/// Read a server log of the RC line by line into LogFile
FUNCTION_BLOCK MC_ReadServerLogFB EXTENDS RobotLibraryBaseExecuteFB
// -------------------------------------------------------------------------
//  SRCI Robot Library
// -------------------------------------------------------------------------
//
//  Object:      MC_ReadServerLogFB
//  Author:      Thorsten Brach
//  Date:        2026-10-23
//
//  Description:
//    ReadServerLog (spec 6.2.6, type 9004): reads the server log ParCmd.ServerLogID from
//    ParCmd.StartLine on into the array LogFile, one CSV line per element. The RC sends a log line in
//    parts of up to 179 characters; the block joins them. The transfer ends with Done when the RC
//    reports the end of the log or when LogFile is full. A rising edge of Execute during the transfer
//    starts it again.
//    Telegram layout of SRCI SDK 1.1.2 (Offset as request counter, IsStartOfLine / IsEndOfLine /
//    EndOfLogReached / LogLine in the response); spec table 6-123 / 6-124 differ.
//
//  Copyright:
//    (C) 2026 Thorsten Brach. All rights reserved
//             Licensed under the MIT License.
//
//  Disclaimer:
//    This project is provided without any guarantee and can be used for
//    private and commercial purposes. Any use is at the user's
//    own risk and responsibility.
//
// -------------------------------------------------------------------------
VAR_INPUT
  /// command parameter
  ParCmd          : ReadServerLogParCmd;
END_VAR
VAR_OUTPUT
  /// Command is transferred and confirmed by the RC
  CommandBuffered : BOOL;
  /// command outputs
  OutCmd          : ReadServerLogOutCmd;
END_VAR
VAR_IN_OUT
  /// Requested log file: one log line per element
  LogFile         : ARRAY [*] OF STRING(RobotLibraryParameter.LOG_LINE_LEN);
END_VAR
VAR
  /// internal copy of command parameter
 _parCmd          : ReadServerLogParCmd;
  /// command data to send
 _command         : ReadServerLogSendData;
  /// response data received
 _response        : ReadServerLogRecvData;
  /// a part of the log was received and must be stored in LogFile (StoreLogContent)
 _contentReceived : BOOL;
  /// the response to the current Offset was handled
 _offsetHandled   : BOOL;
  /// new rising edge of Execute during the transfer: start again after the end of this one
 _restart         : BOOL;
  /// index of the element of LogFile for the current log line
 _line            : DINT;
  /// number of elements of LogFile used by this transfer
 _lines           : DINT;
  /// a log line is open (parts received, end of line not yet)
 _lineOpen        : BOOL;
  /// characters of the current log line
 _lineLen         : DINT;
  /// characters copied from the received part
 _copyLen         : DINT;
END_VAR

            SUPER^(AxesGroup := AxesGroup);

// store the received part of the log (LogFile is only reachable in the call of the block)
StoreLogContent( AxesGroup := AxesGroup, LogFile := LogFile );
          

METHOD INTERNAL CheckAddParameter : BOOL
VAR_INPUT
  /// Payload pointer
  PayloadPtr : UDINT;
END_VAR
VAR
  /// Payload as byte array
  Payload    : ARRAY [1..SIZEOF(_command)] OF BYTE;
  /// Null Byte array
  Null       : ARRAY [1..SIZEOF(_command)] OF BYTE;
  /// Data length to compare
  DataLen    : UDINT;
END_VAR
                  // Payload pointer must be decreased by one byte, because ADR(Payload) is already one byte !
PayloadPtr := LIMIT (0, PayloadPtr - 1, SIZEOF(Payload) -1);
// Convert command struct to payload array
SysDepMemCpy( pDest := ADR(Payload), pSrc := ADR(_command), DataLen := SIZEOF(_command));
// Calculate the data length to compare - at least one byte must be compared !
DataLen := LIMIT(1, SIZEOF(Payload) - PayloadPtr, SIZEOF(Payload));
// Compare Payload-Array with Null-Byte-Array
CheckAddParameter := SysDepMemCmp( pData1 := ADR(Payload) + PayloadPtr , pData2 := ADR(Null), DataLen := DataLen) <>  RobotLibraryConstants.OK ;
                
END_METHOD

METHOD PROTECTED CheckFunctionSupported : BOOL
VAR_IN_OUT
  /// Robot assignment of function
  AxesGroup : AxesGroup;
END_VAR
                  // ReadServerLog is a mandatory function of the profile Core (spec table 6-119): the RC
// reports no bit for it in RCSupportedFunctions
CheckFunctionSupported := TRUE;
                
END_METHOD

METHOD PROTECTED CheckParameterChanged : BOOL
VAR_IN_OUT
  /// Robot assignment of function
  AxesGroup    : AxesGroup;
END_VAR
                  // The parameters of the transfer are taken with the rising edge of Execute; during the transfer
// only the block itself sends updates (next part of the log: Offset, end: Enable FALSE)
IF ( _stepCmd = 0 )
THEN
  RETURN;
END_IF

IF ( _parameterUpdateInternal )
THEN
  // reset internal flag for send parameter update
 _parameterUpdateInternal := FALSE;
  // inc parameter sequence
 _command.ParSeq := _command.ParSeq + 1;
  // update command data
  CommandData := CreateCommandPayload(AxesGroup := AxesGroup); // ( Access via reference to rCommandFB in ACR )
  // notify active command register
  AxesGroup.Acyclic.ActiveCommandRegister.NotifyParameterChanged := _uniqueID;
END_IF
                
END_METHOD

METHOD PROTECTED CheckParameterValid : BOOL
VAR_IN_OUT
  /// Robot assignment of function
  AxesGroup : AxesGroup;
END_VAR
                  CheckParameterValid := TRUE;

// Check ParCmd.ExportMode: only 0 (output LogFile), the export to a file is optional (table 6-119)
IF ( ParCmd.ExportMode <> 0 )
THEN
  // Parameter not valid
  CheckParameterValid := FALSE;
  // Set error
  SetError( ErrorID := RobotLibraryErrorIdEnum.ERR_EXPORTMODE_NOT_EXIST, Overwrite := TRUE );
  // Create log entry
  CreateLogMessagePara1 ( Timestamp   := AxesGroup.State.SystemTime,
                          MessageType := MessageType.CMD,
                          Severity    := Severity.ERROR,
                          MessageCode := ErrorID,
                          MessageText := 'Invalid Parameter ParCmd.ExportMode = {1}',
                          Para1       := USINT_TO_STRING(ParCmd.ExportMode));
  RETURN;
END_IF

// Check ParCmd.StartLine: the first line is 1 (log header)
IF ( ParCmd.StartLine = 0 )
THEN
  // Parameter not valid
  CheckParameterValid := FALSE;
  // Set error
  SetError( ErrorID := RobotLibraryErrorIdEnum.ERR_INVALID_PAR_CMD, Overwrite := TRUE );
  // Create log entry
  CreateLogMessagePara1 ( Timestamp   := AxesGroup.State.SystemTime,
                          MessageType := MessageType.CMD,
                          Severity    := Severity.ERROR,
                          MessageCode := ErrorID,
                          MessageText := 'Invalid Parameter ParCmd.StartLine = {1}',
                          Para1       := UDINT_TO_STRING(ParCmd.StartLine));
  RETURN;
END_IF

// Check ParCmd.ServerLogID: -1 (latest), 0 (oldest) or an ID
IF ( ParCmd.ServerLogID < -1 )
THEN
  // Parameter not valid
  CheckParameterValid := FALSE;
  // Set error
  SetError( ErrorID := RobotLibraryErrorIdEnum.ERR_INVALID_PAR_CMD, Overwrite := TRUE );
  // Create log entry
  CreateLogMessagePara1 ( Timestamp   := AxesGroup.State.SystemTime,
                          MessageType := MessageType.CMD,
                          Severity    := Severity.ERROR,
                          MessageCode := ErrorID,
                          MessageText := 'Invalid Parameter ParCmd.ServerLogID = {1}',
                          Para1       := INT_TO_STRING(ParCmd.ServerLogID));
  RETURN;
END_IF
                
END_METHOD

METHOD INTERNAL CreateCommandPayload : RobotLibraryCommandDataFB
VAR_IN_OUT
  /// Robot assignment of function
  AxesGroup : AxesGroup;
END_VAR
VAR
  /// internal index for loops
 _idx          : DINT;
  /// Parameter count
 _parameterCnt : DINT;
END_VAR
// Sent CMD payload (PLC to RC) of "ReadServerLog" - layout of SRCI SDK 1.1.2 (spec table 6-123
// has no Offset, ContextFilter at byte 12)
// --------------------------
// Header
// --------------------------
// Byte 00 : UINT  - Type HB
// Byte 01 :       - Type LB
// Byte 02 : USINT - Reserve | ExecutionMode
// Byte 03 : USINT - ParSeq  | Priority
// --------------------------
// Datablock
// --------------------------
// Byte 04 : BYTE  - Bit 0: Enable
// Byte 05 : BYTE  - Reserved
// Byte 06 : UINT  - ServerLogID HB
// Byte 07 :       - ServerLogID LB
// Byte 08 : UDINT - StartLine
// Byte 12 : UDINT - Offset
// Byte 16 : USINT - ContextFilter[0]
// ...
// Byte 25 : USINT - ContextFilter[9]
// --------------------------
                  // set command parameter
_command.CmdTyp      :=  CmdType.ReadServerLog;
// spec table 6-121: parallel only (default of ExecMode, FB_init)
_command.ExecMode    :=  ExecMode;
_command.ParSeq      := _command.ParSeq;
_command.Priority    :=  Priority;
_command.Reserve     := 0;
// -1 (latest) -> 16#FFFF
_command.ServerLogID := INT_TO_UINT(_parCmd.ServerLogID);
_command.StartLine   := _parCmd.StartLine;
FOR _idx := 0 TO 9
DO
  _command.ContextFilter[_idx] := _parCmd.ContextFilter[_idx];
END_FOR

// copy command data to header
_cmdHeader := _command;
// call base implementation to copy header to payload buffer
CreateCommandPayload := SUPER^.CreateCommandPayload(AxesGroup := AxesGroup);

// Check parameter must be added ?
IF ( CheckAddParameter(CreateCommandPayload.PayloadPtr))
THEN
  // add command.Enable
  CreateCommandPayload.AddBool(_command.Enable);
  // inc parameter counter
 _parameterCnt := _parameterCnt + 1;
END_IF

// Check parameter must be added ?
IF ( CheckAddParameter(CreateCommandPayload.PayloadPtr))
THEN
  // add command.Reserve
  CreateCommandPayload.AddByte(_command.Reserve);
  // inc parameter counter
 _parameterCnt := _parameterCnt + 1;
END_IF

// Check parameter must be added ?
IF ( CheckAddParameter(CreateCommandPayload.PayloadPtr))
THEN
  // add command.ServerLogID
  CreateCommandPayload.AddUint(_command.ServerLogID);
  // inc parameter counter
 _parameterCnt := _parameterCnt + 1;
END_IF

// Check parameter must be added ?
IF ( CheckAddParameter(CreateCommandPayload.PayloadPtr))
THEN
  // add command.StartLine
  CreateCommandPayload.AddUdint(_command.StartLine);
  // inc parameter counter
 _parameterCnt := _parameterCnt + 1;
END_IF

// Check parameter must be added ?
IF ( CheckAddParameter(CreateCommandPayload.PayloadPtr))
THEN
  // add command.Offset
  CreateCommandPayload.AddUdint(_command.Offset);
  // inc parameter counter
 _parameterCnt := _parameterCnt + 1;
END_IF

FOR _idx := 0 TO 9
DO
  // Check parameter must be added ?
  IF ( CheckAddParameter(CreateCommandPayload.PayloadPtr))
  THEN
    // add command.ContextFilter[x]
    CreateCommandPayload.AddUsint(_command.ContextFilter[_idx]);
    // inc parameter counter
   _parameterCnt := _parameterCnt + 1;
  END_IF
END_FOR

// Create logging
CreateCommandPayloadLog(AxesGroup := AxesGroup, ParameterCnt := _parameterCnt);
                
END_METHOD

METHOD INTERNAL CreateCommandPayloadLog
VAR_IN_OUT
  /// Robot assignment of function
  AxesGroup : AxesGroup;
END_VAR
VAR_INPUT
  /// Parameter count
  ParameterCnt : DINT;
END_VAR
VAR
  /// internal index for loops
 _idx : DINT;
END_VAR
                  // Create log entry for Parameter start
CreateLogMessagePara1 ( Timestamp   := AxesGroup.State.SystemTime,
                        MessageType := MessageType.CMD,
                        Severity    := Severity.DEBUG,
                        MessageCode := 0,
                        MessageText := 'Create command payload with {1} parameter(s) :',
                        Para1       := DINT_TO_STRING(ParameterCnt));

// Return if no parameter is remaining...
IF ( ParameterCnt = 0 ) THEN RETURN; END_IF
// dec remaining parameter(s)
ParameterCnt := ParameterCnt - 1;
// Create log entry for Command.Enable
CreateLogMessagePara1 ( Timestamp   := AxesGroup.State.SystemTime,
                        MessageType := MessageType.CMD,
                        Severity    := Severity.DEBUG,
                        MessageCode := 0,
                        MessageText := 'Command.Enable = {1}',
                        Para1       :=  BOOL_TO_STRING(_command.Enable));

// Return if no parameter is remaining...
IF ( ParameterCnt = 0 ) THEN RETURN; END_IF
// dec remaining parameter(s)
ParameterCnt := ParameterCnt - 1;
// Create log entry for Command.Reserve
CreateLogMessagePara1 ( Timestamp   := AxesGroup.State.SystemTime,
                        MessageType := MessageType.CMD,
                        Severity    := Severity.DEBUG,
                        MessageCode := 0,
                        MessageText := 'Command.Reserve = {1}',
                        Para1       :=  BYTE_TO_STRING(_command.Reserve));

// Return if no parameter is remaining...
IF ( ParameterCnt = 0 ) THEN RETURN; END_IF
// dec remaining parameter(s)
ParameterCnt := ParameterCnt - 1;
// Create log entry for Command.ServerLogID
CreateLogMessagePara1 ( Timestamp   := AxesGroup.State.SystemTime,
                        MessageType := MessageType.CMD,
                        Severity    := Severity.DEBUG,
                        MessageCode := 0,
                        MessageText := 'Command.ServerLogID = {1}',
                        Para1       :=  UINT_TO_STRING(_command.ServerLogID));

// Return if no parameter is remaining...
IF ( ParameterCnt = 0 ) THEN RETURN; END_IF
// dec remaining parameter(s)
ParameterCnt := ParameterCnt - 1;
// Create log entry for Command.StartLine
CreateLogMessagePara1 ( Timestamp   := AxesGroup.State.SystemTime,
                        MessageType := MessageType.CMD,
                        Severity    := Severity.DEBUG,
                        MessageCode := 0,
                        MessageText := 'Command.StartLine = {1}',
                        Para1       :=  UDINT_TO_STRING(_command.StartLine));

// Return if no parameter is remaining...
IF ( ParameterCnt = 0 ) THEN RETURN; END_IF
// dec remaining parameter(s)
ParameterCnt := ParameterCnt - 1;
// Create log entry for Command.Offset
CreateLogMessagePara1 ( Timestamp   := AxesGroup.State.SystemTime,
                        MessageType := MessageType.CMD,
                        Severity    := Severity.DEBUG,
                        MessageCode := 0,
                        MessageText := 'Command.Offset = {1}',
                        Para1       :=  UDINT_TO_STRING(_command.Offset));

FOR _idx := 0 TO 9
DO
  // Return if no parameter is remaining...
  IF ( ParameterCnt = 0 ) THEN RETURN; END_IF
  // dec remaining parameter(s)
  ParameterCnt := ParameterCnt - 1;
  // Create log entry for Command.ContextFilter
  CreateLogMessagePara2 ( Timestamp   := AxesGroup.State.SystemTime,
                          MessageType := MessageType.CMD,
                          Severity    := Severity.DEBUG,
                          MessageCode := 0,
                          MessageText := 'Command.ContextFilter[{2}] = {1}',
                          Para1       :=  USINT_TO_STRING(_command.ContextFilter[_idx]),
                          Para2       :=  DINT_TO_STRING(_idx));
END_FOR
                
END_METHOD

METHOD FB_init : BOOL
VAR_INPUT
  /// if TRUE, the retain variables are initialized (warm start / cold start)
  bInitRetains : BOOL;
  /// if TRUE, the instance afterwards gets moved into the copy code (online change)
  bInCopyCode  : BOOL;
END_VAR
                  MyType := 'MC_ReadServerLogFB';

// spec 6.2.6: processed with low priority because of its processing time
ExecMode := ExecutionMode.PARALLEL;
Priority := PriorityLevel.LOW;
                
END_METHOD

METHOD PROTECTED OnApplyOutCmd
VAR_INPUT
  /// Command message state
  State : CmdMessageState;
END_VAR
                  IF ( State = CmdMessageState.EMPTY )
THEN
  // Reset command outputs
  SysDepMemSet(pDest := ADR(OutCmd), Value := 0, DataLen := SIZEOF(OutCmd));
END_IF

// the counters of the log come with every part (StoreLogContent), the received lines are counted there
                
END_METHOD

METHOD PROTECTED OnExecRun : DINT
VAR_IN_OUT
  /// Robot assignment of function
  AxesGroup : AxesGroup;
END_VAR
                  // call base implementation
SUPER^.OnExecRun(AxesGroup := AxesGroup);

CASE _stepCmd OF

  00:  IF (( _execute_R.Q ) OR ( _restart )) AND ( NOT Error )
       THEN
        _restart := FALSE;
         // Check function is supported and parameter are valid ?
         IF (( CheckFunctionSupported( AxesGroup := AxesGroup )) AND
             ( CheckParameterValid   ( AxesGroup := AxesGroup )))
         THEN
           // set busy flag
           Busy := TRUE;
           // Reset command outputs
           SysDepMemSet(pDest := ADR(OutCmd), Value := 0, DataLen := SIZEOF(OutCmd));
           // apply command parameter
          _parCmd := ParCmd;
           // first element of LogFile, no open line
          _line            := 0;
          _lines           := 0;
          _lineOpen        := FALSE;
          _lineLen         := 0;
          _contentReceived := FALSE;
          _offsetHandled   := FALSE;
           // transfer on, first request
          _command.Enable := TRUE;
          _command.Offset := 1;
           // init parameter sequence
          _command.ParSeq := 1;
           // create command data
           CommandData := CreateCommandPayload(AxesGroup := AxesGroup);
           // Add command to active command register
          _uniqueID := AxesGroup.Acyclic.ActiveCommandRegister.AddCmd( pCommandFB := ADR(THIS^ ));
           // set timeout
           SetTimeout(PT := _timeoutCmd, rTimer := _timerCmd);
           // inc step counter
          _stepCmd := _stepCmd + 1;
         END_IF
       END_IF

  01:  // spec 6.2.6: a new rising edge of Execute during the transfer aborts it and starts the
       // command again. SRCI SDK 1.1 keeps the read position of a running command, so the transfer
       // ends first (Enable FALSE) and the command is added again (new ACR entry).
       IF ( _executeRestart_R.Q ) AND ( NOT _restart )
       THEN
        _restart := TRUE;
        _command.Enable := FALSE;
        _parameterUpdateInternal := TRUE;
       END_IF

       // Wait for responce received
       IF ( _responseReceived )
       THEN
         // reset response received flag
        _responseReceived := FALSE;

         CASE _response.State OF
           CmdMessageState.DONE:
             IF ( _restart )
             THEN
               // the old transfer ended: start again (step 00)
               Reset();
              _restart := TRUE;
             ELSE
               OnUpdateStateFlags(_response.State);
               // set timeout
               SetTimeout(PT := _timeoutCmd, rTimer := _timerCmd);
               // inc step counter
              _stepCmd := _stepCmd + 1;
             END_IF

           CmdMessageState.ABORTED, CmdMessageState.ERROR:
            _restart := FALSE;
             OnUpdateStateFlags(_response.State);
             // set timeout
             SetTimeout(PT := _timeoutCmd, rTimer := _timerCmd);
             // inc step counter
            _stepCmd := _stepCmd + 1;

         ELSE
           OnUpdateStateFlags(_response.State);
           // a part of the log for the current request ? (responses to older requests are ignored)
           IF (( _command.Enable                     ) AND
               ( NOT _restart                        ) AND
               ( NOT _offsetHandled                  ) AND
               ( _response.Offset = _command.Offset  ))
           THEN
            _offsetHandled   := TRUE;
            _contentReceived := TRUE;
           END_IF
         END_CASE
       END_IF

  02: IF ( NOT Execute)
      THEN
        Reset();
      END_IF

ELSE
  // invalid step
  SetError( ErrorID := RobotLibraryErrorIdEnum.ERR_INVALID_STEP, Overwrite := TRUE );
END_CASE

// Reset FB
IF ( NOT Execute ) AND ( NOT _restart )
THEN
  Reset();
END_IF
                
END_METHOD

METHOD PROTECTED OnUpdateStateFlags
VAR_INPUT
  /// Command message state
  State : CmdMessageState;
END_VAR
                  // Reset State flags
Done := FALSE;

CASE State OF
  // No operation or process is active
  CmdMessageState.EMPTY               :;
  // Created but not yet started
  CmdMessageState.CREATED             :;
  // Buffered and awaiting execution
  CmdMessageState.BUFFERED            : CommandBuffered := TRUE;
  // Buffered in planner for future execution
  CmdMessageState.BUFFERED_IN_PLANNER : CommandBuffered := TRUE;
  // Currently active and in progress
  CmdMessageState.ACTIVE              : CommandBuffered := TRUE;
  // Interrupted and awaiting continuation
  CmdMessageState.INTERRUPTED         :;
  // Requested for abort
  CmdMessageState.ABORT_REQUEST       :;
  // Successfully completed
  CmdMessageState.DONE                : Done            := TRUE;
                                        Busy            := FALSE;
  // Aborted before completion
  CmdMessageState.ABORTED             : Busy            := FALSE;
  // Encountered an error during execution
  CmdMessageState.ERROR               : Error           := TRUE;
                                        Busy            := FALSE;
END_CASE
                
END_METHOD

METHOD INTERNAL ParseResponsePayload : DINT
VAR_INPUT
  /// Response data
  ResponseData : RobotLibraryResponseDataFB;
  /// Timestamp
  Timestamp    : SystemTime;
END_VAR
VAR
  /// Parameter count
 _parameterCnt : DINT;
  /// Byte 13: line flags
 _flags        : BYTE;
END_VAR
// Received CMD payload (RC to PLC) of "ReadServerLog" - layout of SRCI SDK 1.1.2 (spec table
// 6-124: byte 13 only IsSplitLine, LogContent from byte 14)
// --------------------------
// Header
// --------------------------
// Byte 00 : USINT   - ParSeq | State
// Byte 01 : SINT    - AlarmMessageSeverity
// Byte 02 : UINT    - AlarmMessageCode HB
// Byte 03 :         - AlarmMessageCode LB
// --------------------------
// Datablock
// --------------------------
// Byte 04 : UDINT   - AvailableLogLines
// Byte 08 : UDINT   - AvailableFilteredLogLines
// Byte 12 : USINT   - LogContentLength
// Byte 13 : BYTE    - Bit 0: IsStartOfLine, Bit 1: IsEndOfLine, Bit 2: EndOfLogReached
// Byte 14 : UDINT   - LogLine
// Byte 18 : UDINT   - Offset
// Byte 22 : CHAR    - LogContent[0]
// ...
// Byte 200: CHAR    - LogContent[178]
// --------------------------
                  // call base implementation to parse the header from payload buffer
ResponseData.PayloadPtr := SUPER^.ParseResponsePayload(ResponseData := ResponseData, Timestamp := Timestamp);

// missing (trailing zero) bytes of the payload are 0, no values of the previous response
SysDepMemSet( pDest := ADR(_response), Value := 0, DataLen := SIZEOF(_response));

// copy parsed header to response
_response.ParSeq               := _rspHeader.ParSeq;
_response.State                := _rspHeader.State;
_response.AlarmMessageSeverity := _rspHeader.AlarmMessageSeverity;
_response.AlarmMessageCode     := _rspHeader.AlarmMessageCode;

// Check payload remaining ?
IF ( ResponseData.IsPayloadRemaining)
THEN
  // Get Response.AvailableLogLines
 _response.AvailableLogLines := ResponseData.GetUdint();
  // inc parameter counter
 _parameterCnt := _parameterCnt + 1;
END_IF

// Check payload remaining ?
IF ( ResponseData.IsPayloadRemaining)
THEN
  // Get Response.AvailableFilteredLogLines
 _response.AvailableFilteredLogLines := ResponseData.GetUdint();
  // inc parameter counter
 _parameterCnt := _parameterCnt + 1;
END_IF

// Check payload remaining ?
IF ( ResponseData.IsPayloadRemaining)
THEN
  // Get Response.LogContentLength
 _response.LogContentLength := ResponseData.GetUsint();
  // inc parameter counter
 _parameterCnt := _parameterCnt + 1;
END_IF

// Check payload remaining ?
IF ( ResponseData.IsPayloadRemaining)
THEN
  // Get Response.IsStartOfLine / IsEndOfLine / EndOfLogReached
 _flags                     := ResponseData.GetByte();
 _response.IsStartOfLine    := _flags.0;
 _response.IsEndOfLine      := _flags.1;
 _response.EndOfLogReached  := _flags.2;
  // inc parameter counter
 _parameterCnt := _parameterCnt + 1;
END_IF

// Check payload remaining ?
IF ( ResponseData.IsPayloadRemaining)
THEN
  // Get Response.LogLine
 _response.LogLine := ResponseData.GetUdint();
  // inc parameter counter
 _parameterCnt := _parameterCnt + 1;
END_IF

// Check payload remaining ?
IF ( ResponseData.IsPayloadRemaining)
THEN
  // Get Response.Offset
 _response.Offset := ResponseData.GetUdint();
  // inc parameter counter
 _parameterCnt := _parameterCnt + 1;
END_IF

// Check payload remaining ?
IF ( ResponseData.IsPayloadRemaining ) AND ( _response.LogContentLength > 0 )
THEN
  // Get Response.LogContent (LogContentLength characters)
 _response.LogContent := ResponseData.GetString( Size := MIN( USINT_TO_DINT(_response.LogContentLength), RobotLibraryConstants.SERVER_LOG_CONTENT_MAX ));
  // inc parameter counter
 _parameterCnt := _parameterCnt + 1;
END_IF

// Create logging
ParseResponsePayloadLog(ResponseData := ResponseData, Timestamp := Timestamp, ParameterCnt := _parameterCnt);
                
END_METHOD

METHOD INTERNAL ParseResponsePayloadLog
VAR_INPUT
  /// Response data
  ResponseData : RobotLibraryResponseDataFB;
  /// Timestamp
  Timestamp    : SystemTime;
  /// Parameter count
  ParameterCnt : DINT;
END_VAR
                  // Create log entry for Parameter start
CreateLogMessagePara1 ( Timestamp   := Timestamp,
                        MessageType := MessageType.CMD,
                        Severity    := Severity.DEBUG,
                        MessageCode := 0,
                        MessageText := '{1} parameter(s) to parse from the response data:',
                        Para1       := DINT_TO_STRING(ParameterCnt));

// Return if no parameter is remaining...
IF ( ParameterCnt = 0 ) THEN RETURN; END_IF
// dec remaining parameter(s)
ParameterCnt := ParameterCnt - 1;
// Create log entry for AvailableLogLines
CreateLogMessagePara1 ( Timestamp   := Timestamp,
                        MessageType := MessageType.CMD,
                        Severity    := Severity.DEBUG,
                        MessageCode := 0,
                        MessageText := 'Response.AvailableLogLines = {1}',
                        Para1       :=  UDINT_TO_STRING(_response.AvailableLogLines));

// Return if no parameter is remaining...
IF ( ParameterCnt = 0 ) THEN RETURN; END_IF
// dec remaining parameter(s)
ParameterCnt := ParameterCnt - 1;
// Create log entry for AvailableFilteredLogLines
CreateLogMessagePara1 ( Timestamp   := Timestamp,
                        MessageType := MessageType.CMD,
                        Severity    := Severity.DEBUG,
                        MessageCode := 0,
                        MessageText := 'Response.AvailableFilteredLogLines = {1}',
                        Para1       :=  UDINT_TO_STRING(_response.AvailableFilteredLogLines));

// Return if no parameter is remaining...
IF ( ParameterCnt = 0 ) THEN RETURN; END_IF
// dec remaining parameter(s)
ParameterCnt := ParameterCnt - 1;
// Create log entry for LogContentLength
CreateLogMessagePara1 ( Timestamp   := Timestamp,
                        MessageType := MessageType.CMD,
                        Severity    := Severity.DEBUG,
                        MessageCode := 0,
                        MessageText := 'Response.LogContentLength = {1}',
                        Para1       :=  USINT_TO_STRING(_response.LogContentLength));

// Return if no parameter is remaining...
IF ( ParameterCnt = 0 ) THEN RETURN; END_IF
// dec remaining parameter(s)
ParameterCnt := ParameterCnt - 1;
// Create log entry for IsStartOfLine
CreateLogMessagePara1 ( Timestamp   := Timestamp,
                        MessageType := MessageType.CMD,
                        Severity    := Severity.DEBUG,
                        MessageCode := 0,
                        MessageText := 'Response.IsStartOfLine = {1}',
                        Para1       :=  BOOL_TO_STRING(_response.IsStartOfLine));

// Return if no parameter is remaining...
IF ( ParameterCnt = 0 ) THEN RETURN; END_IF
// dec remaining parameter(s)
ParameterCnt := ParameterCnt - 1;
// Create log entry for LogLine
CreateLogMessagePara1 ( Timestamp   := Timestamp,
                        MessageType := MessageType.CMD,
                        Severity    := Severity.DEBUG,
                        MessageCode := 0,
                        MessageText := 'Response.LogLine = {1}',
                        Para1       :=  UDINT_TO_STRING(_response.LogLine));

// Return if no parameter is remaining...
IF ( ParameterCnt = 0 ) THEN RETURN; END_IF
// dec remaining parameter(s)
ParameterCnt := ParameterCnt - 1;
// Create log entry for Offset
CreateLogMessagePara1 ( Timestamp   := Timestamp,
                        MessageType := MessageType.CMD,
                        Severity    := Severity.DEBUG,
                        MessageCode := 0,
                        MessageText := 'Response.Offset = {1}',
                        Para1       :=  UDINT_TO_STRING(_response.Offset));

// Return if no parameter is remaining...
IF ( ParameterCnt = 0 ) THEN RETURN; END_IF
// dec remaining parameter(s)
ParameterCnt := ParameterCnt - 1;
// Create log entry for LogContent
CreateLogMessagePara1 ( Timestamp   := Timestamp,
                        MessageType := MessageType.CMD,
                        Severity    := Severity.DEBUG,
                        MessageCode := 0,
                        MessageText := 'Response.LogContent = {1}',
                        Para1       :=  _response.LogContent);
                
END_METHOD

METHOD PROTECTED Reset : DINT
VAR_INPUT
END_VAR
                  Reset := SUPER^.Reset();

Done             := FALSE;
Busy             := FALSE;
CommandBuffered  := FALSE;
_restart         := FALSE;
_contentReceived := FALSE;
_offsetHandled   := FALSE;
_command.Enable  := FALSE;
                
END_METHOD

METHOD PRIVATE StoreLogContent
VAR_IN_OUT
  /// Robot assignment of function
  AxesGroup : AxesGroup;
  /// Requested log file: one log line per element
  LogFile : ARRAY [*] OF STRING(RobotLibraryParameter.LOG_LINE_LEN);
END_VAR
VAR
  /// LogFile is full
  Full : BOOL;
END_VAR
                  IF ( NOT _contentReceived )
THEN
  RETURN;
END_IF
_contentReceived := FALSE;

OutCmd.AvailableLogLines         := _response.AvailableLogLines;
OutCmd.AvailableFilteredLogLines := _response.AvailableFilteredLogLines;

// a part of a log line ? (a response without log line: the RC had not read the log yet)
IF ( _response.LogLine > 0 ) AND (( _response.LogContentLength > 0 ) OR ( _response.IsEndOfLine ))
THEN
  // a new line starts in the next element of LogFile
  IF (( _response.IsStartOfLine ) OR ( NOT _lineOpen ))
  THEN
   _line  := LOWER_BOUND(LogFile, 1) + _lines;
   _lines := _lines + 1;
    SysDepMemSet( pDest := ADR(LogFile[_line]), Value := 0, DataLen := SIZEOF(LogFile[_line]) );
   _lineLen  := 0;
   _lineOpen := TRUE;
  END_IF

  // append the part (a line longer than LOG_LINE_LEN is cut)
 _copyLen := MIN( USINT_TO_DINT(_response.LogContentLength), RobotLibraryParameter.LOG_LINE_LEN - _lineLen );
  IF ( _copyLen > 0 )
  THEN
    SysDepMemCpy( pDest := ADR(LogFile[_line]) + _lineLen, pSrc := ADR(_response.LogContent), DataLen := DINT_TO_UDINT(_copyLen) );
   _lineLen := _lineLen + _copyLen;
  ELSIF ( _response.LogContentLength > 0 )
  THEN
    CreateLogMessagePara1 ( Timestamp   := AxesGroup.State.SystemTime,
                            MessageType := MessageType.CMD,
                            Severity    := Severity.WARNING,
                            MessageCode := 0,
                            MessageText := 'Log line {1} longer than LOG_LINE_LEN, cut',
                            Para1       := UDINT_TO_STRING(_response.LogLine));
  END_IF

  IF ( _response.IsEndOfLine )
  THEN
   _lineOpen               := FALSE;
    OutCmd.ReceivedLogLines := OutCmd.ReceivedLogLines + 1;
    OutCmd.LogLine          := _response.LogLine;
    IF ( _response.AvailableFilteredLogLines > 0 )
    THEN
      OutCmd.Progress := MIN( 100.0, UDINT_TO_REAL(OutCmd.ReceivedLogLines) * 100.0 / UDINT_TO_REAL(_response.AvailableFilteredLogLines) );
    END_IF
  END_IF
END_IF

OutCmd.EndOfLogReached := _response.EndOfLogReached;
// no element of LogFile left for another line
Full := ( NOT _lineOpen ) AND ( LOWER_BOUND(LogFile, 1) + _lines > UPPER_BOUND(LogFile, 1) );

IF (( _response.EndOfLogReached ) OR ( Full ))
THEN
  // end of the transfer: Enable FALSE, the RC answers with DONE
 _command.Enable := FALSE;
ELSE
  // next part of the log
 _command.Offset := _command.Offset + 1;
 _offsetHandled  := FALSE;
END_IF
_parameterUpdateInternal := TRUE;
                
END_METHOD
END_FUNCTION_BLOCK

FUNCTION_BLOCK MC_ReadServerLog EXTENDS RobotLibraryBaseFB
VAR
END_VAR

            
          

METHOD FB_init : BOOL
VAR_INPUT
  /// if TRUE, the retain variables are initialized (warm start / cold start)
  bInitRetains : BOOL; 
  /// if TRUE, the instance afterwards gets moved into the copy code (online change)
  bInCopyCode  : BOOL;  
END_VAR
                  MyType := 'MC_ReadServerLogFB';

ExecMode := ExecutionMode.PARALLEL;
Priority := PriorityLevel.NORMAL;
                
END_METHOD
END_FUNCTION_BLOCK

/// Restart/reboot of the RC.
FUNCTION_BLOCK MC_RestartControllerFB EXTENDS RobotLibraryBaseExecuteFB
// ------------------------------------------------------------------------- 
//  SRCI Robot Library                                                
// ------------------------------------------------------------------------- 
//                                                                           
//  Object:      RestartControllerFB                                       
//  Author:      Thorsten Brach                                                
//  Date:        2024-06-01
//
//  Description:                                              
//   
//                                                                           
//  Copyright: 
//    (C) 2024 Thorsten Brach. All rights reserved                                                                                                                                            
//             Licensed under the MIT License.
//                                                                           
//  Disclaimer:                                                                           
//    This project is provided without any guarantee and can be used for   
//    private and commercial purposes. Any use is at the user’s 
//    own risk and responsibility.
//
// -------------------------------------------------------------------------
VAR_INPUT
  /// Command parameter 
  ParCmd          : RestartControllerParCmd;  
END_VAR

VAR_OUTPUT
  /// Command is transferred and confirmed by the RC
  CommandBuffered : BOOL;
  /// Command outputs 
  OutCmd          : RestartControllerOutCmd;  
END_VAR

VAR
  /// internal copy of command parameter 
 _parCmd          : RestartControllerParCmd;
  /// command data to send
 _command         : RestartControllerSendData;
  /// response data received
 _response        : RestartControllerRecvData;      
END_VAR

            SUPER^(AxesGroup := AxesGroup);
          

METHOD INTERNAL CheckAddParameter : BOOL
VAR_INPUT
  /// Payload pointer
  PayloadPtr : UDINT;
END_VAR
VAR
  /// Payload as byte array
  Payload    : ARRAY [1..SIZEOF(_command)] OF BYTE;
  /// Null Byte array 
  Null       : ARRAY [1..SIZEOF(_command)] OF BYTE;
  /// Data length to compare
  DataLen    : UDINT;
END_VAR
                  // Payload pointer must be decreased by one byte, because ADR(Payload) is already one byte !
PayloadPtr := LIMIT (0, PayloadPtr - 1, SIZEOF(Payload) -1);
// Convert command struct to payload array
SysDepMemCpy( pDest := ADR(Payload), pSrc := ADR(_command), DataLen := SIZEOF(_command));
// Calculate the data length to compare - at least one byte must be compared !
DataLen := LIMIT(1, SIZEOF(Payload) - PayloadPtr, SIZEOF(Payload)); 
// Compare Payload-Array with Null-Byte-Array
CheckAddParameter := SysDepMemCmp( pData1 := ADR(Payload) + PayloadPtr , pData2 := ADR(Null), DataLen := DataLen) <>  RobotLibraryConstants.OK ;
                
END_METHOD

METHOD PROTECTED CheckFunctionSupported : BOOL
VAR_IN_OUT
  /// Robot assignment of function
  AxesGroup : AxesGroup; 
END_VAR
                  CheckFunctionSupported := AxesGroup.State.RobotData.RCSupportedFunctions.RestartController;

IF ( NOT CheckFunctionSupported )
THEN
  // call base implementation for set error and create log entry
  SUPER^.CheckFunctionSupported(AxesGroup := AxesGroup);
END_IF
                
END_METHOD

METHOD PROTECTED CheckParameterChanged : BOOL
VAR_IN_OUT
  /// Robot assignment of function
  AxesGroup    : AxesGroup; 
END_VAR
                  // Check ParCmd Size is > 0, because MemCmp does not work correctly with size = 0
IF (SIZEOF(ParCmd) = 0) OR (_stepCmd = 0)
THEN 
  RETURN;
END_IF

// compare memory 
_parameterChanged := ( SysDepMemCmp(pData1 := ADR(ParCmd), pData2 := ADR(_parCmd), DataLen := SIZEOF(ParCmd)) <> RobotLibraryConstants.OK );

// check parameter valid ?
_parameterValid   := CheckParameterValid( AxesGroup := AxesGroup );

IF ((  _parameterChanged        )  AND 
    (  _parameterValid          )) OR
    (  _parameterUpdateInternal )  
THEN  
  // Create log entry for parameter changed event
  CreateLogMessagePara1 ( Timestamp   := AxesGroup.State.SystemTime,
                          MessageType := MessageType.CMD,
                          Severity    := Severity.DEBUG,
                          MessageCode := 0,
                          MessageText := 'NotifyParameterChanged Event {1}',
                          Para1       :=  '' );

  // reset internal flag for send parameter update
 _parameterUpdateInternal := FALSE;
  // update internal copy of parameters 
 _parCmd := ParCmd;
  // inc parameter sequence
 _command.ParSeq := _command.ParSeq + 1;
  // update command data  
  CommandData := CreateCommandPayload(AxesGroup := AxesGroup); // ( Access via reference to rCommandFB in ACR )
  // notify active command register 
  AxesGroup.Acyclic.ActiveCommandRegister.NotifyParameterChanged := _uniqueID;
END_IF
                
END_METHOD

METHOD INTERNAL CreateCommandPayload : RobotLibraryCommandDataFB
VAR_IN_OUT
  /// Robot assignment of function
  AxesGroup : AxesGroup; 
END_VAR
VAR
  /// Parameter count
 _parameterCnt : DINT;
END_VAR
// Table 6-57: Sent CMD payload (PLC to RC) of "RestartController"
// --------------------------
// Header
// --------------------------
// Byte 00 : UINT  - Type HB     
// Byte 01 :       - Type LB    
// Byte 02 : USINT - Reserve | ExecutionMode
// Byte 03 : USINT - ParSeq  | Priority
// --------------------------
                  // set command parameter 
_command.CmdTyp     :=  CmdType.RestartController;
_command.ExecMode   :=  ExecMode;
_command.ParSeq     := _command.ParSeq;
_command.Priority   :=  Priority;


// copy command data to header
_cmdHeader := _command;
// call base implementation to copy header to payload buffer
CreateCommandPayload := SUPER^.CreateCommandPayload(AxesGroup := AxesGroup);


// Create logging
CreateCommandPayloadLog(AxesGroup := AxesGroup, ParameterCnt := _parameterCnt);
                
END_METHOD

METHOD INTERNAL CreateCommandPayloadLog
VAR_IN_OUT
  /// Robot assignment of function
  AxesGroup : AxesGroup; 
END_VAR
VAR_INPUT
  /// Parameter count
  ParameterCnt : DINT;
END_VAR
                  // Create log entry for Parameter start
CreateLogMessagePara1 ( Timestamp   := AxesGroup.State.SystemTime,
                        MessageType := MessageType.CMD,
                        Severity    := Severity.DEBUG,
                        MessageCode := 0,
                        MessageText := 'Create command payload with {1} parameter(s) :',
                        Para1       := DINT_TO_STRING(ParameterCnt));
                
END_METHOD

METHOD FB_init : BOOL
VAR_INPUT
  /// if TRUE, the retain variables are initialized (warm start / cold start)
  bInitRetains : BOOL; 
  /// if TRUE, the instance afterwards gets moved into the copy code (online change)
  bInCopyCode  : BOOL;  
END_VAR
                  MyType := 'MC_RestartControllerFB';

ExecMode := ExecutionMode.PARALLEL;
Priority := PriorityLevel.NORMAL;
                
END_METHOD

METHOD PROTECTED OnApplyOutCmd
VAR_INPUT
  /// Command message state
  State : CmdMessageState;
END_VAR
                  IF ( State = CmdMessageState.EMPTY ) 
THEN
  // Reset command outputs
  SysDepMemSet(pDest := ADR(OutCmd), Value := 0, DataLen := SIZEOF(OutCmd));         
END_IF

IF (( State = CmdMessageState.ACTIVE ) OR
    ( State = CmdMessageState.DONE   ))
THEN
  // Update results
  OutCmd.RestartAccepted := _response.RestartAccepted;
END_IF
                
END_METHOD

METHOD PROTECTED OnExecRun : DINT
VAR_IN_OUT
  /// Robot assignment of function
  AxesGroup : AxesGroup; 
END_VAR
                  // call base implementation
SUPER^.OnExecRun(AxesGroup := AxesGroup);

CASE _stepCmd OF
  
  00:  IF ( _execute_R.Q ) AND ( NOT Error)   
       THEN
         // Check function is supported and parameter are valid ?
         IF (( CheckFunctionSupported( AxesGroup := AxesGroup )) AND
             ( CheckParameterValid   ( AxesGroup := AxesGroup )))      
         THEN
           // set busy flag
           Busy := TRUE;
           // Reset command outputs
           SysDepMemSet(pDest := ADR(OutCmd), Value := 0, DataLen := SIZEOF(OutCmd));         
           // apply command parameter
          _parCmd := ParCmd;
           // init parameter sequence
          _command.ParSeq := 1;
           // create command data
           CommandData := CreateCommandPayload(AxesGroup := AxesGroup);
           // Add command to active command register
          _uniqueID := AxesGroup.Acyclic.ActiveCommandRegister.AddCmd( pCommandFB := ADR(THIS^ ));     
           // set timeout
           SetTimeout(PT := _timeoutCmd, rTimer := _timerCmd);
           // inc step counter
          _stepCmd := _stepCmd + 1;
         END_IF 
       END_IF
     

  01:  // Wait for responce received
       IF ( _responseReceived )
       THEN
         // reset response received flag
        _responseReceived := FALSE;
         // update state flags
         OnUpdateStateFlags(_response.State);
         // update state flags
         OnApplyOutCmd(_response.State);

         // Done, Aborted or Error ?
         IF (_response.State >= CmdMessageState.DONE )
         THEN
           // set timeout
           SetTimeout(PT := _timeoutCmd, rTimer := _timerCmd);
           // inc step counter
          _stepCmd := _stepCmd + 1; 
         END_IF
       END_IF


  02: IF ( NOT Execute)
      THEN
        Reset();
      END_IF     

ELSE
  // invalid step
  SetError( ErrorID := RobotLibraryErrorIdEnum.ERR_INVALID_STEP, Overwrite := TRUE );
END_CASE


// Reset FB
IF ( NOT Execute )
THEN
  Reset();
END_IF
                
END_METHOD

METHOD PROTECTED OnUpdateStateFlags
VAR_INPUT
  /// Command message state
  State : CmdMessageState;
END_VAR
                  // Reset State flags
Done := FALSE;

CASE State OF

  // No operation or process is active
  CmdMessageState.EMPTY               :;
  // Created but not yet started
  CmdMessageState.CREATED             :;
  // Buffered and awaiting execution
  CmdMessageState.BUFFERED            : CommandBuffered    := TRUE;
  // Buffered in planner for future execution
  CmdMessageState.BUFFERED_IN_PLANNER : CommandBuffered    := TRUE;
  // Currently active and in progress
  CmdMessageState.ACTIVE              :;
  // Interrupted and awaiting continuation
  CmdMessageState.INTERRUPTED         :;  
  // Requested for abort
  CmdMessageState.ABORT_REQUEST       :;
  // Successfully completed
  CmdMessageState.DONE                : Done               := TRUE;
                                        Busy               := FALSE;
  // Aborted before completion
  CmdMessageState.ABORTED             : Busy               := FALSE;
  // Encountered an error during execution
  CmdMessageState.ERROR               : Error              := TRUE;
                                        Busy               := FALSE;
END_CASE
                
END_METHOD

METHOD INTERNAL ParseResponsePayload : DINT
VAR_INPUT
  /// Response data
  ResponseData : RobotLibraryResponseDataFB;
  /// Timestamp
  Timestamp    : SystemTime;  
END_VAR
VAR
  /// Parameter count
 _parameterCnt : DINT;
END_VAR
// Table 6-58: Received CMD payload (RC to PLC) of "RestartController"
// --------------------------
// Header
// --------------------------
// Byte 00 : USINT - ParSeq | State     
// Byte 01 : SINT  - AlarmMessageSeverity    
// Byte 02 : UINT  - AlarmMessageCode HB
// Byte 03 :       - AlarmMessageCode LB
// --------------------------
// Datablock
// --------------------------
// Byte 4  : BOOL  - RestartAccepted
                  // call base implementation to parse the header from payload buffer
ResponseData.PayloadPtr := SUPER^.ParseResponsePayload(ResponseData := ResponseData, Timestamp := Timestamp);

// ST-FIX F100: missing (trailing zero) bytes of the payload are 0, no values of the previous response
SysDepMemSet( pDest := ADR(_response), Value := 0, DataLen := SIZEOF(_response));

// copy parsed header to response
_response.ParSeq               := _rspHeader.ParSeq;
_response.State                := _rspHeader.State;
_response.AlarmMessageSeverity := _rspHeader.AlarmMessageSeverity;
_response.AlarmMessageCode     := _rspHeader.AlarmMessageCode;

// Check payload remaining ? 
IF ( ResponseData.IsPayloadRemaining)
THEN 
  // Get Response.RestartAccepted
 _response.RestartAccepted := ResponseData.GetBool();
  // inc parameter counter
 _parameterCnt := _parameterCnt + 1;
END_IF


// Create logging
ParseResponsePayloadLog(ResponseData := ResponseData, Timestamp := Timestamp, ParameterCnt := _parameterCnt);
                
END_METHOD

METHOD INTERNAL ParseResponsePayloadLog
VAR_INPUT
  /// Response data
  ResponseData : RobotLibraryResponseDataFB;
  /// Timestamp
  Timestamp    : SystemTime;  
  /// Parameter count
  ParameterCnt : DINT;
END_VAR
                  // Create log entry for Parameter start
CreateLogMessagePara1 ( Timestamp   := Timestamp,
                        MessageType := MessageType.CMD,
                        Severity    := Severity.DEBUG,
                        MessageCode := 0,
                        MessageText := '{1} parameter(s) to parse from the response data:',
                        Para1       := DINT_TO_STRING(ParameterCnt));
                        

// Return if no parameter is remaining...
IF ( ParameterCnt = 0 ) THEN RETURN; END_IF
// dec remaining parameter(s)                        
ParameterCnt := ParameterCnt - 1;
// Create log entry for RestartAccepted
CreateLogMessagePara1 ( Timestamp   := Timestamp,
                        MessageType := MessageType.CMD,
                        Severity    := Severity.DEBUG,
                        MessageCode := 0,
                        MessageText := 'Response.RestartAccepted = {1}',
                        Para1       :=  BOOL_TO_STRING(_response.RestartAccepted));


                
END_METHOD

METHOD PROTECTED Reset : DINT
VAR_INPUT
END_VAR
                  Reset := SUPER^.Reset();

Done               := FALSE;
Busy               := FALSE;
CommandBuffered    := FALSE;

                
END_METHOD
END_FUNCTION_BLOCK

/// Handles multiple mechanisms required for operation of the interface.
/// For maximal performance, this FB must be called after the function FB's, 
/// so that the data can be written to the fieldbus in the same cycle as the start of FB occours 
FUNCTION_BLOCK MC_RobotTaskFB EXTENDS RobotLibraryLogFB
// ------------------------------------------------------------------------- 
//  SRCI Robot Library                                                
// ------------------------------------------------------------------------- 
//                                                                           
//  Object:      RobotTaskFB                                       
//  Author:      Thorsten Brach                                                
//  Date:        2024-06-01
//
//  Description:                                              
//   
//                                                                           
//  Copyright: 
//    (C) 2024 Thorsten Brach. All rights reserved                                                                                                                                            
//             Licensed under the MIT License.
//                                                                           
//  Disclaimer:                                                                           
//    This project is provided without any guarantee and can be used for   
//    private and commercial purposes. Any use is at the user’s 
//    own risk and responsibility.
//
// -------------------------------------------------------------------------
VAR_INPUT
  /// Set TRUE (default) to initialize the interface
  Enable            : BOOL;
  /// User defined robot name
  RobotName         : STRING(20);
  /// Current System Time
  SystemTime        : SystemTime;
  /// Online Change detected
  OnlineChange      : BOOL;
  /// Axes Group ID -> is used to uniquely identify each RA on a per RC basis.
  ///
  /// The IDs start with 0: an RC with only one RA uses ID 0.
  /// ST-FIX F138: spec V1.5.9 says 1 (one RA) and 1-15 (several RAs); this is an error of the spec
  /// (confirmed by PI), the SDK uses 0 too.
  AxesGroupID       : BYTE := 0;
  /// Configuration parameter
  ParCfg            : RobotTaskParCfg;
END_VAR

VAR_IN_OUT
  /// Inputs of PLC for communication from RC
  RobotInData       : ARRAY[*] OF BYTE;
  /// Outputs of PLC for communication to RC
  RobotOutData      : ARRAY[*] OF BYTE;
  ///  User data stored on the PLC according to Table 6-10
  UserData          : UserData;
  /// ToolData stored on PLC. For more information refer to 5.5.6.3
  ToolData          : ARRAY[*] OF Tool;
  /// LoadData stored on PLC.For more information refer to 5.5.6.4
  FrameData         : ARRAY[*] OF Frame;
  /// LoadData stored on PLC.For more information refer to 5.5.6.4 
  LoadData          : ARRAY[*] OF Load;
  /// Work areas stored on PLC. For more information refer to 5.5.8
  WorkAreas         : ARRAY[*] OF RobotWorkArea;
  /// Software limits stored on PLC
  SWLimits          : SWLimits;
  /// Default dynamics stored on PLC. For more information refer to 5.5.7
  DefaultDynamics   : DefaultDynamics;
  /// Reference dynamics stored on PLC. For more information refer to 5.5.7
  ReferenceDynamics : ReferenceDynamics;
  /// System log on PLC
  SystemLog         : ARRAY[0..RobotLibraryParameter.SYSTEM_LOG_MAX ] OF STRING(RobotLibraryParameter.MESSAGE_TEXT_LEN);
  /// Message buffer on the PLC - For more information refer to 5.5.11
  MessageLog        : ARRAY[0..RobotLibraryParameter.MESSAGE_LOG_MAX] OF AlarmMessage;
  /// Robot assignment of function
  AxesGroup         : AxesGroup;
END_VAR

VAR_OUTPUT
  /// FB is being processed
  Busy              : BOOL;
  /// Interface is initialized (RI state: "Initialized").
  /// For more information on RI states refer to chapter 5.5.3.1.
  Initialized       : BOOL;
  /// Server and client were successfully synchronized (RI state: "Synchronized").
  /// For more information on the synchronization mechanism refer to chapter 5.6.7.
  Synchronized      : BOOL;
  /// An error occurred
  Error             : BOOL;
  /// ErrorID reported by RC for error identification according to Table 7-1
  ErrorID           : WORD;
  ErrorIdEnum       : RobotLibraryErrorIdEnum;  
  ErrorAddTxt       : STRING(RobotLibraryConstants.MAX_ADD_TEXT_LENGTH);
  /// WarningID for warning identification reported during execution of command according to Table 7-3
  WarningID         : WORD;
  WarningIdEnum     : RobotLibraryWarningIdEnum;  
  /// InfoID for info identification reported during execution of command according to Table 7-5
  InfoID            : WORD;    
  InfoIdEnum        : RobotLibraryInfoIdEnum;    
END_VAR

VAR
  /// internal copy of configuration parameter
 _parCfg                       : RobotTaskParCfg;

  /// internal ToolData for comparation to user ToolData
 _toolData                     : ARRAY[0..RobotLibraryParameter.TOOL_MAX       -1] OF Tool;
  /// internal FrameData for comparation to user FrameData
 _frameData                    : ARRAY[0..RobotLibraryParameter.FRAME_MAX      -1] OF Frame;
  /// internal LoadData for comparation to user LoadData
 _loadData                     : ARRAY[0..RobotLibraryParameter.LOAD_MAX       -1] OF Load;
  /// internal WorkAreas for comparation to user WorkAreas
 _workAreas                    : ARRAY[0..RobotLibraryParameter.WORK_AREAS_MAX -1] OF RobotWorkArea;
  /// internal Software limits for comparation to user Software limit
 _swLimits                     : SWLimits;
  /// internal default dynamics for comparation to user default dynamics
 _defaultDynamics              : DefaultDynamics;
  /// internal reference dynamics for comparation to user reference dynamics
 _referenceDynamics            : ReferenceDynamics;

  /// FB for exchange configuration
 _exchangeConfiguration        : MC_ExchangeConfigurationFB;
  /// FB for read robot data
 _readRobotData                : MC_ReadRobotDataFB;
  /// FB for read messaged
 _readMessages                 : MC_ReadMessagesFB;  
  /// FB for read tool data
 _readToolData                 : MC_ReadToolDataFB;  
  /// FB for read frame data
 _readFrameData                : MC_ReadFrameDataFB;  
  /// FB for read load data
 _readLoadData                 : MC_ReadLoadDataFB;  
  /// FB for read work area
 _readWorkArea                 : MC_ReadWorkAreaFB;  
  /// FB for read robot software limits
 _readRobotSWLimits            : MC_ReadRobotSWLimitsFB;  
  /// FB for read robot default dynamics
 _readRobotDefaultDynamics     : MC_ReadRobotDefaultDynamicsFB;  
  /// FB for read robot reference dynamics
 _readRobotReferenceDynamics   : MC_ReadRobotReferenceDynamicsFB;  

  /// FB for write tool data
 _writeToolData                : MC_WriteToolDataFB;  
  /// FB for write frame data
 _writeFrameData               : MC_WriteFrameDataFB;  
  /// FB for write load data
 _writeLoadData                : MC_WriteLoadDataFB;  
  /// FB for write work area
 _writeWorkArea                : MC_WriteWorkAreaFB;  
  /// FB for write robot software limits
 _writeRobotSWLimits           : MC_WriteRobotSWLimitsFB;  
  /// FB for write robot default dynamics
 _writeRobotDefaultDynamics    : MC_WriteRobotDefaultDynamicsFB;  
  /// FB for write robot reference dynamics
 _writeRobotReferenceDynamics  : MC_WriteRobotReferenceDynamicsFB;  
  /// Send Buffer
  SendData                     : RobotLibrarySendDataFB;
  /// Recv Buffer
  RecvData                     : RobotLibraryRecvDataFB;
  /// Telegram 
  Telegram                     : Telegram; 
  
  /// internal step counter for command
 _stepCmd                      : DINT;
  /// internal timer for command 
  {attribute 'hide'}
 _timerCmd                     : TON;
  /// internal timeout for command
  {attribute 'hide'}
 _timeoutCmd                   : TIME := T#5S; 

  /// internal step counter for synchronisation of frame data
 _stepSyncFrameData            : DINT;
  /// internal timer for synchronisation of frame data
  {attribute 'hide'}
 _timerSyncFrameData           : TON;
  /// internal timeout for synchronisation of frame data
  {attribute 'hide'}
 _timeoutSyncFrameData         : TIME := T#5S;
   /// internal index for frame data synchronisation
 _syncIdxFrameData             : USINT;
  /// internal index for maximal amount of frames data( MIN(PLC,RC) ) 
 _syncIdxMaxFrameData          : DINT;
 
  /// internal step counter for synchronisation of load data
 _stepSyncLoadData             : DINT;
  /// internal timer for synchronisation of load data
  {attribute 'hide'}
 _timerSyncLoadData             : TON;
  /// internal timeout for synchronisation of load data
  {attribute 'hide'}
 _timeoutSyncLoadData           : TIME := T#5S; 
  /// internal index for load data synchronisation
 _syncIdxLoadData               : USINT;
  /// internal index for maximal amount of load data ( MIN(PLC,RC) ) 
 _syncIdxMaxLoadData            : DINT;

  /// internal step counter for synchronisation of tool data
 _stepSyncToolData              : DINT;
  /// internal timer for synchronisation of tool data
  {attribute 'hide'}
 _timerSyncToolData             : TON;
  /// internal timeout for synchronisation of tool data
  {attribute 'hide'}
 _timeoutSyncToolData           : TIME := T#5S; 
  /// internal index for tool data synchronisation
 _syncIdxToolData               : USINT;
  /// internal index for maximal amount of tool data ( MIN(PLC,RC) ) 
 _syncIdxMaxToolData            : DINT;

  /// internal step counter for synchronisation of work areas
 _stepSyncWorkArea            : DINT;
 /// internal timer for synchronisation of work areas
  {attribute 'hide'}
 _timerSyncWorkArea           : TON;
  /// internal timeout for synchronisation of work areas
  {attribute 'hide'}
 _timeoutSyncWorkArea         : TIME := T#5S; 
  /// internal index for WorkArea synchronisation
 _syncIdxWorkArea             : USINT;
  /// internal index for maximal amount of Work Area( MIN(PLC,RC) ) 
 _syncIdxMaxWorkArea          : DINT;
 
  /// internal step counter for synchronisation of software limits
 _stepSyncSWLimits            : DINT;
  /// internal timer for synchronisation of software limits
  {attribute 'hide'}
 _timerSyncSWLimits           : TON;
  /// internal timeout for synchronisation of software limits
  {attribute 'hide'}
 _timeoutSyncSWLimits         : TIME := T#5S; 

  /// internal step counter for synchronisation of default dynamics
 _stepSyncDefaultDynamics      : DINT;
  /// internal timer for synchronisation of default dynamics
  {attribute 'hide'}
 _timerSyncDefaultDynamics     : TON;
  /// internal timeout for synchronisation of default dynamics
  {attribute 'hide'}
 _timeoutSyncDefaultDynamics   : TIME := T#5S; 
 
  /// internal step counter for synchronisation of reference dynamics
 _stepSyncReferenceDynamics    : DINT;
  /// internal timer for synchronisation of reference dynamics
  {attribute 'hide'}
 _timerSyncReferenceDynamics   : TON;
  /// internal timeout for synchronisation of reference dynamics
  {attribute 'hide'}
 _timeoutSyncReferenceDynamics : TIME := T#5S; 


 
 
  /// Rising edge for enable
  {attribute 'hide'}
 _enable_R                    : R_TRIG;
  /// Falling edge for enable
  {attribute 'hide'}
 _enable_F                    : F_TRIG;

  /// Flag that indicated the the connection is alive (data exchange)
 _aliveBit                    : BOOL;
  /// last lifesign counter value
 _aliveValue                  : BYTE;
  /// timer for detecting alive state
 _aliveCheck                  : TON;
  /// rising edge for connection is alive
  {attribute 'hide'}
 _alive_R                     : R_TRIG;
  /// falling edge for connection is alive
  {attribute 'hide'}
 _alive_F                     : F_TRIG;
   /// last telegram state
 _lastTelegramState           : TelegramState   := TelegramState.UNDEFINED;
   /// last telegram control
 _lastTelegramControl         : ControlHalfByte := ControlHalfByte.NONE;
END_VAR

VAR // CONSTANT
  /// Lower array dimension of RobotInData
  ROBOT_IN_DATA_MIN   : DINT;
  /// Upper array dimension of RobotInData
  ROBOT_IN_DATA_MAX   : DINT;
  /// Size of RobotInData
  ROBOT_IN_DATA_SIZE  : UDINT;
  /// Lower array dimension of RobotOutData
  ROBOT_OUT_DATA_MIN  : DINT;
  /// Upper array dimension of RobotOutData
  ROBOT_OUT_DATA_MAX  : DINT;
  /// Size of RobotOutData
  ROBOT_OUT_DATA_SIZE : UDINT;
END_VAR

VAR CONSTANT
  {attribute 'hide'}
  FRAGMENT_HEADER_SIZE : UDINT := SIZEOF(TelegramPlcToRobFragmentHeader);
  /// Size of the comand header
  {attribute 'hide'}
  COMMAND_HEADER_SIZE  : UDINT := SIZEOF(TelegramPlcToRobCommandHeader);
  /// Size of the footer
  {attribute 'hide'}
  FOOTER_SIZE          : UDINT := 1;
  /// Minimal payload size for telegram
  {attribute 'hide'}
  MIN_PAYLOAD_SIZE     : UDINT := 1;
  /// Active command
  {attribute 'hide'}
  ACTIVE_CMD           : UDINT := 1;
  /// Buffered command
  {attribute 'hide'}
  BUFFER_CMD           : UDINT := 2;
  /// Empty command entry
  {attribute 'hide'}
  EMPTY_CMD_ENTRY      : AxesGroupAcyclicAcrEntryCmdBuffer := (State := BufferStateCmd.EMPTY);
  /// bitmask to mask the LifeSign out of the halfbyte
  {attribute 'hide'}
  LIFESIGN_BIT_MASK    : BYTE := 2#000_1111;   
  /// Primary sequence
  {attribute 'hide'}
  PRIMARY_SEQUENCE     : DINT := 0;
  /// Secondary sequence
  {attribute 'hide'}
  SECONDARY_SEQUENCE   : DINT := 1;  
  /// Empty Execution-Order-List entry
  {attribute 'hide'}
  EMPTY_EOL_ENTRY      : DINT := 0;
END_VAR
            
          
VAR
  /// ST-FIX F63: telegram sequence that is handled/filled first (lower Seq/Ack number)
  _seqSendFirst : DINT;
  /// ST-FIX F63: loop counter over the telegram sequences in Seq order
  _seqOrderIdx : DINT;
  /// ST-FIX F63: distance of two Seq numbers
  _seqDiff : DINT;
  /// ST-FIX F63: next Seq number
  _seqNext : UINT;
END_VAR

VAR
  /// ST-FIX F65: telegram sequence timeout (4 x LifeSignTimeOut without new Seq number)
  _seqAckTimeout : TON;
  /// ST-FIX F66: lifesign of header and footer differ -> frame is not processed
  _frameInvalid : BOOL;
  /// ST-FIX F79: last error state of the RC during the initialization (reported at the init timeout)
  _initErrorState : TelegramState;
END_VAR

VAR
  _turns : BYTE; // ST-FIX F60: turn number nibble
END_VAR

VAR
  _restartReset : BOOL; // ST-FIX F23: interface reset on the RC requested by a restart
END_VAR

VAR
  /// ST-FIX F132: identification of this instance (1..n, assigned in FB_init, kept by an online change)
 _instanceId : UDINT;
END_VAR

VAR_STAT
  /// ST-FIX F132: number of RobotTask instances created (source of _instanceId)
 _instanceCount   : UDINT;
  /// ST-FIX F132: instance that uses the telegram buffers of the entry (0 = free entry)
 _peripheryOwner  : ARRAY[1..PERIPHERY_ENTRIES] OF UDINT;
  /// ST-FIX F132: address of RobotInData of the entry
 _peripheryInAdr  : ARRAY[1..PERIPHERY_ENTRIES] OF PVOID;
  /// ST-FIX F132: address of RobotOutData of the entry
 _peripheryOutAdr : ARRAY[1..PERIPHERY_ENTRIES] OF PVOID;
END_VAR

VAR CONSTANT
  /// ST-FIX F132: number of RobotTask instances whose telegram buffers are checked
  PERIPHERY_ENTRIES : DINT := 16;
END_VAR

            // Get array dimension of RobotInData
ROBOT_IN_DATA_MIN  := LOWER_BOUND  ( RobotInData,1);
ROBOT_IN_DATA_MAX  := UPPER_BOUND  ( RobotInData,1);
ROBOT_IN_DATA_SIZE := DINT_TO_UDINT( ROBOT_IN_DATA_MAX - ROBOT_IN_DATA_MIN + 1);

// Get array dimension of RobotInData
ROBOT_OUT_DATA_MIN  := LOWER_BOUND  ( RobotOutData,1);
ROBOT_OUT_DATA_MAX  := UPPER_BOUND  ( RobotOutData,1);
ROBOT_OUT_DATA_SIZE := DINT_TO_UDINT( ROBOT_OUT_DATA_MAX - ROBOT_OUT_DATA_MIN + 1);

// ST-FIX F132: an AxesGroup and the telegram buffers belong to one RobotTask only (table 7-1:
// 16#8007 / 16#8008); a second instance does nothing else, so it cannot disturb the first one
IF ( NOT CheckAssignmentValid( AxesGroup    := AxesGroup,
                               RobotInData  := RobotInData,
                               RobotOutData := RobotOutData ) )
THEN
  Error       := HasError;
  ErrorIdEnum := ErrorID;
  RETURN;
END_IF

HandleAxesGroup              ( AxesGroup         := AxesGroup,
	                             ToolData          := ToolData, 
	                             FrameData         := FrameData, 
	                             LoadData          := LoadData, 
	                             WorkAreas         := WorkAreas, 
	                             SWLimits          := SWLimits, 
	                             DefaultDynamics   := DefaultDynamics, 
	                             ReferenceDynamics := ReferenceDynamics);
                               
HandleLifeSign               ( AxesGroup         := AxesGroup);
HandleLogMessagesAck         ( AxesGroup         := AxesGroup);
HandleInvalidFrames          ( AxesGroup         := AxesGroup, RobotInData := RobotInData);
HandleTelegramStateCtrl      (                               );
HandleAliveBit               ( RobotInData[1]                );
HandleSeqAck                 ( AxesGroup         := AxesGroup);
HandleUserData               ( AxesGroup         := AxesGroup, UserData := UserData );

HandleSync                   ( AxesGroup         := AxesGroup,
                               ToolData          := ToolData,
                               FrameData         := FrameData,
                               LoadData          := LoadData,
                               WorkAreas         := WorkAreas,
                               SWLimits          := SWLimits,
                               DefaultDynamics   := DefaultDynamics,
                               ReferenceDynamics := ReferenceDynamics);

OnCall                       ( AxesGroup         := AxesGroup);
OnExecRun                    ( AxesGroup         := AxesGroup);

AxesGroupToTelegram          ( AxesGroup         := AxesGroup );

CreateSendPayload            ( AxesGroup         := AxesGroup, RobotOutData := RobotOutData );
IF ( NOT _frameInvalid ) // ST-FIX F66
THEN
  ParseRecvPayload             ( AxesGroup         := AxesGroup, RobotInData  := RobotInData);
END_IF 

AxesGroupFromTelegram        ( AxesGroup         := AxesGroup);


// call internal functionblocks
_exchangeConfiguration      ( Name := RobotName, ExecMode := ExecutionMode.PARALLEL, Priority := PriorityLevel.NORMAL, AxesGroup := AxesGroup );
_readRobotData              ( Name := RobotName, ExecMode := ExecutionMode.PARALLEL, Priority := PriorityLevel.NORMAL, AxesGroup := AxesGroup );
_readMessages               ( Name := RobotName, ExecMode := ExecutionMode.PARALLEL, Priority := PriorityLevel.NORMAL, AxesGroup := AxesGroup );
_readToolData               ( UpdateSystemData := FALSE, // ST-FIX F16
 Name := RobotName, ExecMode := ExecutionMode.PARALLEL, Priority := PriorityLevel.NORMAL, AxesGroup := AxesGroup );
_readFrameData              ( UpdateSystemData := FALSE, // ST-FIX F16
 Name := RobotName, ExecMode := ExecutionMode.PARALLEL, Priority := PriorityLevel.NORMAL, AxesGroup := AxesGroup );
_readLoadData               ( UpdateSystemData := FALSE, // ST-FIX F16
 Name := RobotName, ExecMode := ExecutionMode.PARALLEL, Priority := PriorityLevel.NORMAL, AxesGroup := AxesGroup );
_readWorkArea               ( UpdateSystemData := FALSE, // ST-FIX F16
 Name := RobotName, ExecMode := ExecutionMode.PARALLEL, Priority := PriorityLevel.NORMAL, AxesGroup := AxesGroup );  
_readRobotSWLimits          ( UpdateSystemData := FALSE, // ST-FIX F16
 Name := RobotName, ExecMode := ExecutionMode.PARALLEL, Priority := PriorityLevel.NORMAL, AxesGroup := AxesGroup );  
_readRobotDefaultDynamics   ( UpdateSystemData := FALSE, // ST-FIX F16
 Name := RobotName, ExecMode := ExecutionMode.PARALLEL, Priority := PriorityLevel.NORMAL, AxesGroup := AxesGroup );
_readRobotReferenceDynamics ( UpdateSystemData := FALSE, // ST-FIX F16
 Name := RobotName, ExecMode := ExecutionMode.PARALLEL, Priority := PriorityLevel.NORMAL, AxesGroup := AxesGroup );
_writeToolData              ( Name := RobotName, ExecMode := ExecutionMode.PARALLEL, Priority := PriorityLevel.NORMAL, AxesGroup := AxesGroup );  
_writeFrameData             ( Name := RobotName, ExecMode := ExecutionMode.PARALLEL, Priority := PriorityLevel.NORMAL, AxesGroup := AxesGroup );  
_writeLoadData              ( Name := RobotName, ExecMode := ExecutionMode.PARALLEL, Priority := PriorityLevel.NORMAL, AxesGroup := AxesGroup );  
_writeWorkArea              ( Name := RobotName, ExecMode := ExecutionMode.PARALLEL, Priority := PriorityLevel.NORMAL, AxesGroup := AxesGroup );  
_writeRobotSWLimits         ( Name := RobotName, ExecMode := ExecutionMode.PARALLEL, Priority := PriorityLevel.NORMAL, AxesGroup := AxesGroup );  
_writeRobotDefaultDynamics  ( Name := RobotName, ExecMode := ExecutionMode.PARALLEL, Priority := PriorityLevel.NORMAL, AxesGroup := AxesGroup );  
_writeRobotReferenceDynamics( Name := RobotName, ExecMode := ExecutionMode.PARALLEL, Priority := PriorityLevel.NORMAL, AxesGroup := AxesGroup );  


// Update SystemLog and MessageLog
SystemLog  := AxesGroup.MessageLog.SystemLogs;
MessageLog := AxesGroup.MessageLog.Messages;
          

METHOD PRIVATE AxesGroupFromTelegram
VAR_IN_OUT
  /// Robot assignment of function
  AxesGroup    : AxesGroup;
END_VAR
                  AxesGroupFromTelegramCyclic         (AxesGroup := AxesGroup);
AxesGroupFromTelegramCyclicOptional (AxesGroup := AxesGroup);
                
END_METHOD

METHOD PRIVATE AxesGroupFromTelegramCyclic
VAR_IN_OUT
  /// Robot assignment of function
  AxesGroup : AxesGroup;
END_VAR
                  // ---------------------------------
// Mapp Telegramm to AxesGroup Data  
// ---------------------------------
AxesGroup.Cyclic.RobToPlc.SRCIVersion    := Telegram.RobToPlc.Header.SRCIVersion ;
AxesGroup.Cyclic.RobToPlc.LifeSign       := Telegram.RobToPlc.Header.LifeSign ;
AxesGroup.Cyclic.RobToPlc.TelegramState  := Telegram.RobToPlc.Header.TelegramState ;
AxesGroup.Cyclic.RobToPlc.StatusRobotArm := DwordToRaStatusWord(Telegram.RobToPlc.Header.StatusRobotArm);
AxesGroup.Cyclic.RobToPlc.Override       := Telegram.RobToPlc.Header.Override ;
                
END_METHOD

METHOD PRIVATE AxesGroupFromTelegramCyclicOptional
VAR_IN_OUT
  /// Robot assignment of function
  AxesGroup: AxesGroup;
END_VAR
                  // Sub ProgramData {{{
AxesGroup.CyclicOptional.RobToPlc.SubProgramData.Data := Telegram.RobToPlc.CyclicOptional.SubProgramData.Data;
// }}}


// Cartesian position {{{
AxesGroup.CyclicOptional.RobToPlc.CartesianPosition.Active                   :=                                     AxesGroup.CyclicOptional.RobToPlc.CartesianPosition.Active;
AxesGroup.CyclicOptional.RobToPlc.CartesianPosition.X                        :=                                      Telegram.RobToPlc.CyclicOptional.CartesianPosition.X;
AxesGroup.CyclicOptional.RobToPlc.CartesianPosition.Y                        :=                                      Telegram.RobToPlc.CyclicOptional.CartesianPosition.Y;
AxesGroup.CyclicOptional.RobToPlc.CartesianPosition.Z                        :=                                      Telegram.RobToPlc.CyclicOptional.CartesianPosition.Z;
AxesGroup.CyclicOptional.RobToPlc.CartesianPosition.Rx                       :=                                      Telegram.RobToPlc.CyclicOptional.CartesianPosition.Rx;
AxesGroup.CyclicOptional.RobToPlc.CartesianPosition.Ry                       :=                                      Telegram.RobToPlc.CyclicOptional.CartesianPosition.Ry;
AxesGroup.CyclicOptional.RobToPlc.CartesianPosition.Rz                       :=                                      Telegram.RobToPlc.CyclicOptional.CartesianPosition.Rz;
AxesGroup.CyclicOptional.RobToPlc.CartesianPosition.Config.Shoulder          :=              WordToArmConfigShoulder(Telegram.RobToPlc.CyclicOptional.CartesianPosition.Config);
AxesGroup.CyclicOptional.RobToPlc.CartesianPosition.Config.Elbow             :=              WordToArmConfigElbow   (Telegram.RobToPlc.CyclicOptional.CartesianPosition.Config);
AxesGroup.CyclicOptional.RobToPlc.CartesianPosition.Config.Wrist             :=              WordToArmConfigWrist   (Telegram.RobToPlc.CyclicOptional.CartesianPosition.Config);
_turns := GetHalfeByteLo(Telegram.RobToPlc.CyclicOptional.CartesianPosition.Turns_J2_J1); // ST-FIX F60: sign + magnitude (spec 5.5.4.4)
AxesGroup.CyclicOptional.RobToPlc.CartesianPosition.TurnNumber.J1Turns := BYTE_TO_SINT(_turns AND 16#07);
IF ( ( _turns AND 16#08 ) <> 0 )
THEN
  AxesGroup.CyclicOptional.RobToPlc.CartesianPosition.TurnNumber.J1Turns := INT_TO_SINT(-SINT_TO_INT(AxesGroup.CyclicOptional.RobToPlc.CartesianPosition.TurnNumber.J1Turns));
END_IF
_turns := GetHalfeByteHi(Telegram.RobToPlc.CyclicOptional.CartesianPosition.Turns_J2_J1); // ST-FIX F60: sign + magnitude (spec 5.5.4.4)
AxesGroup.CyclicOptional.RobToPlc.CartesianPosition.TurnNumber.J2Turns := BYTE_TO_SINT(_turns AND 16#07);
IF ( ( _turns AND 16#08 ) <> 0 )
THEN
  AxesGroup.CyclicOptional.RobToPlc.CartesianPosition.TurnNumber.J2Turns := INT_TO_SINT(-SINT_TO_INT(AxesGroup.CyclicOptional.RobToPlc.CartesianPosition.TurnNumber.J2Turns));
END_IF
_turns := GetHalfeByteLo(Telegram.RobToPlc.CyclicOptional.CartesianPosition.Turns_J4_J3); // ST-FIX F60: sign + magnitude (spec 5.5.4.4)
AxesGroup.CyclicOptional.RobToPlc.CartesianPosition.TurnNumber.J3Turns := BYTE_TO_SINT(_turns AND 16#07);
IF ( ( _turns AND 16#08 ) <> 0 )
THEN
  AxesGroup.CyclicOptional.RobToPlc.CartesianPosition.TurnNumber.J3Turns := INT_TO_SINT(-SINT_TO_INT(AxesGroup.CyclicOptional.RobToPlc.CartesianPosition.TurnNumber.J3Turns));
END_IF
_turns := GetHalfeByteHi(Telegram.RobToPlc.CyclicOptional.CartesianPosition.Turns_J4_J3); // ST-FIX F60: sign + magnitude (spec 5.5.4.4)
AxesGroup.CyclicOptional.RobToPlc.CartesianPosition.TurnNumber.J4Turns := BYTE_TO_SINT(_turns AND 16#07);
IF ( ( _turns AND 16#08 ) <> 0 )
THEN
  AxesGroup.CyclicOptional.RobToPlc.CartesianPosition.TurnNumber.J4Turns := INT_TO_SINT(-SINT_TO_INT(AxesGroup.CyclicOptional.RobToPlc.CartesianPosition.TurnNumber.J4Turns));
END_IF
_turns := GetHalfeByteLo(Telegram.RobToPlc.CyclicOptional.CartesianPosition.Turns_J6_J5); // ST-FIX F60: sign + magnitude (spec 5.5.4.4)
AxesGroup.CyclicOptional.RobToPlc.CartesianPosition.TurnNumber.J5Turns := BYTE_TO_SINT(_turns AND 16#07);
IF ( ( _turns AND 16#08 ) <> 0 )
THEN
  AxesGroup.CyclicOptional.RobToPlc.CartesianPosition.TurnNumber.J5Turns := INT_TO_SINT(-SINT_TO_INT(AxesGroup.CyclicOptional.RobToPlc.CartesianPosition.TurnNumber.J5Turns));
END_IF
_turns := GetHalfeByteHi(Telegram.RobToPlc.CyclicOptional.CartesianPosition.Turns_J6_J5); // ST-FIX F60: sign + magnitude (spec 5.5.4.4)
AxesGroup.CyclicOptional.RobToPlc.CartesianPosition.TurnNumber.J6Turns := BYTE_TO_SINT(_turns AND 16#07);
IF ( ( _turns AND 16#08 ) <> 0 )
THEN
  AxesGroup.CyclicOptional.RobToPlc.CartesianPosition.TurnNumber.J6Turns := INT_TO_SINT(-SINT_TO_INT(AxesGroup.CyclicOptional.RobToPlc.CartesianPosition.TurnNumber.J6Turns));
END_IF
AxesGroup.CyclicOptional.RobToPlc.CartesianPosition.TurnNumber.E1Turns := BYTE_TO_SINT(Telegram.RobToPlc.CyclicOptional.CartesianPosition.Turns_E1 AND 16#7F); // ST-FIX F60: sign + magnitude (spec 5.5.4.4)
IF ( ( Telegram.RobToPlc.CyclicOptional.CartesianPosition.Turns_E1 AND 16#80 ) <> 0 )
THEN
  AxesGroup.CyclicOptional.RobToPlc.CartesianPosition.TurnNumber.E1Turns := INT_TO_SINT(-SINT_TO_INT(AxesGroup.CyclicOptional.RobToPlc.CartesianPosition.TurnNumber.E1Turns));
END_IF
AxesGroup.CyclicOptional.RobToPlc.CartesianPosition.E1                       :=                                      Telegram.RobToPlc.CyclicOptional.CartesianPosition.E1;
AxesGroup.CyclicOptional.RobToPlc.CartesianPosition.CoordinateSystem.ToolNo  :=                                      Telegram.RobToPlc.CyclicOptional.CartesianPosition.ToolNo; // ST-FIX F59: tool/frame of the returned position
AxesGroup.CyclicOptional.RobToPlc.CartesianPosition.CurrentCoordinateSystem.ToolNo  :=                                      Telegram.RobToPlc.CyclicOptional.CartesianPosition.CurrentlyUsedToolNo;
AxesGroup.CyclicOptional.RobToPlc.CartesianPosition.CoordinateSystem.FrameNo :=                                      Telegram.RobToPlc.CyclicOptional.CartesianPosition.FrameNo; // ST-FIX F59: tool/frame of the returned position
AxesGroup.CyclicOptional.RobToPlc.CartesianPosition.CurrentCoordinateSystem.FrameNo :=                                      Telegram.RobToPlc.CyclicOptional.CartesianPosition.CurrentlyUsedFrameNo;
// }}}


// Joint position {{{
AxesGroup.CyclicOptional.RobToPlc.JointPosition.Active := AxesGroup.CyclicOptional.RobToPlc.JointPosition.Active;
AxesGroup.CyclicOptional.RobToPlc.JointPosition.J1     :=  Telegram.RobToPlc.CyclicOptional.JointPosition.J1;
AxesGroup.CyclicOptional.RobToPlc.JointPosition.J2     :=  Telegram.RobToPlc.CyclicOptional.JointPosition.J2;
AxesGroup.CyclicOptional.RobToPlc.JointPosition.J3     :=  Telegram.RobToPlc.CyclicOptional.JointPosition.J3;
AxesGroup.CyclicOptional.RobToPlc.JointPosition.J4     :=  Telegram.RobToPlc.CyclicOptional.JointPosition.J4;
AxesGroup.CyclicOptional.RobToPlc.JointPosition.J5     :=  Telegram.RobToPlc.CyclicOptional.JointPosition.J5;
AxesGroup.CyclicOptional.RobToPlc.JointPosition.J6     :=  Telegram.RobToPlc.CyclicOptional.JointPosition.J6;
AxesGroup.CyclicOptional.RobToPlc.JointPosition.E1     :=  Telegram.RobToPlc.CyclicOptional.JointPosition.E1;
// }}}

// Force {{{
AxesGroup.CyclicOptional.RobToPlc.Force.Active          := AxesGroup.CyclicOptional.RobToPlc.Force.Active;
AxesGroup.CyclicOptional.RobToPlc.Force.X               :=  Telegram.RobToPlc.CyclicOptional.Force.X;
AxesGroup.CyclicOptional.RobToPlc.Force.Y               :=  Telegram.RobToPlc.CyclicOptional.Force.Y;
AxesGroup.CyclicOptional.RobToPlc.Force.Z               :=  Telegram.RobToPlc.CyclicOptional.Force.Z;
AxesGroup.CyclicOptional.RobToPlc.Force.Rx              :=  Telegram.RobToPlc.CyclicOptional.Force.Rx;
AxesGroup.CyclicOptional.RobToPlc.Force.Ry              :=  Telegram.RobToPlc.CyclicOptional.Force.Ry;
AxesGroup.CyclicOptional.RobToPlc.Force.Rz              :=  Telegram.RobToPlc.CyclicOptional.Force.Rz;
// }}}

// Current {{{
AxesGroup.CyclicOptional.RobToPlc.Current.Active        := AxesGroup.CyclicOptional.RobToPlc.Current.Active;
AxesGroup.CyclicOptional.RobToPlc.Current.J1            :=  Telegram.RobToPlc.CyclicOptional.Current.J1;
AxesGroup.CyclicOptional.RobToPlc.Current.J2            :=  Telegram.RobToPlc.CyclicOptional.Current.J2;
AxesGroup.CyclicOptional.RobToPlc.Current.J3            :=  Telegram.RobToPlc.CyclicOptional.Current.J3;
AxesGroup.CyclicOptional.RobToPlc.Current.J4            :=  Telegram.RobToPlc.CyclicOptional.Current.J4;
AxesGroup.CyclicOptional.RobToPlc.Current.J5            :=  Telegram.RobToPlc.CyclicOptional.Current.J5;
AxesGroup.CyclicOptional.RobToPlc.Current.J6            :=  Telegram.RobToPlc.CyclicOptional.Current.J6;
// }}}


// Two Sequences {{{
// }}}

// Cartesian Position Extended
AxesGroup.CyclicOptional.RobToPlc.CartesianPositionExt.Active := AxesGroup.CyclicOptional.RobToPlc.CartesianPositionExt.Active;
AxesGroup.CyclicOptional.RobToPlc.CartesianPositionExt.E2     :=  Telegram.RobToPlc.CyclicOptional.CartesianPositionExt.E2;
AxesGroup.CyclicOptional.RobToPlc.CartesianPositionExt.E3     :=  Telegram.RobToPlc.CyclicOptional.CartesianPositionExt.E3;
AxesGroup.CyclicOptional.RobToPlc.CartesianPositionExt.E4     :=  Telegram.RobToPlc.CyclicOptional.CartesianPositionExt.E4;
AxesGroup.CyclicOptional.RobToPlc.CartesianPositionExt.E5     :=  Telegram.RobToPlc.CyclicOptional.CartesianPositionExt.E5;
AxesGroup.CyclicOptional.RobToPlc.CartesianPositionExt.E6     :=  Telegram.RobToPlc.CyclicOptional.CartesianPositionExt.E6;

// Joint Position Extended
AxesGroup.CyclicOptional.RobToPlc.JointPositionExt.Active     := AxesGroup.CyclicOptional.RobToPlc.JointPositionExt.Active;
AxesGroup.CyclicOptional.RobToPlc.JointPositionExt.E2         :=  Telegram.RobToPlc.CyclicOptional.JointPositionExt.E2;
AxesGroup.CyclicOptional.RobToPlc.JointPositionExt.E3         :=  Telegram.RobToPlc.CyclicOptional.JointPositionExt.E3;
AxesGroup.CyclicOptional.RobToPlc.JointPositionExt.E4         :=  Telegram.RobToPlc.CyclicOptional.JointPositionExt.E4;
AxesGroup.CyclicOptional.RobToPlc.JointPositionExt.E5         :=  Telegram.RobToPlc.CyclicOptional.JointPositionExt.E5;
AxesGroup.CyclicOptional.RobToPlc.JointPositionExt.E6         :=  Telegram.RobToPlc.CyclicOptional.JointPositionExt.E6;

// Force Extended
AxesGroup.CyclicOptional.RobToPlc.ForceExt.Active             := AxesGroup.CyclicOptional.RobToPlc.ForceExt.Active;
AxesGroup.CyclicOptional.RobToPlc.ForceExt.E1                 :=  Telegram.RobToPlc.CyclicOptional.ForceExt.E1;
AxesGroup.CyclicOptional.RobToPlc.ForceExt.E2                 :=  Telegram.RobToPlc.CyclicOptional.ForceExt.E2;
AxesGroup.CyclicOptional.RobToPlc.ForceExt.E3                 :=  Telegram.RobToPlc.CyclicOptional.ForceExt.E3;
AxesGroup.CyclicOptional.RobToPlc.ForceExt.E4                 :=  Telegram.RobToPlc.CyclicOptional.ForceExt.E4;
AxesGroup.CyclicOptional.RobToPlc.ForceExt.E5                 :=  Telegram.RobToPlc.CyclicOptional.ForceExt.E5;
AxesGroup.CyclicOptional.RobToPlc.ForceExt.E6                 :=  Telegram.RobToPlc.CyclicOptional.ForceExt.E6;

// Current Extended
AxesGroup.CyclicOptional.RobToPlc.CurrentExt.Active           := AxesGroup.CyclicOptional.RobToPlc.CurrentExt.Active;
AxesGroup.CyclicOptional.RobToPlc.CurrentExt.E1               :=  Telegram.RobToPlc.CyclicOptional.CurrentExt.E1;
AxesGroup.CyclicOptional.RobToPlc.CurrentExt.E2               :=  Telegram.RobToPlc.CyclicOptional.CurrentExt.E2;
AxesGroup.CyclicOptional.RobToPlc.CurrentExt.E3               :=  Telegram.RobToPlc.CyclicOptional.CurrentExt.E3;
AxesGroup.CyclicOptional.RobToPlc.CurrentExt.E4               :=  Telegram.RobToPlc.CyclicOptional.CurrentExt.E4;
AxesGroup.CyclicOptional.RobToPlc.CurrentExt.E5               :=  Telegram.RobToPlc.CyclicOptional.CurrentExt.E5;
AxesGroup.CyclicOptional.RobToPlc.CurrentExt.E6               :=  Telegram.RobToPlc.CyclicOptional.CurrentExt.E6;
                
                
END_METHOD

METHOD PRIVATE AxesGroupToTelegram : DINT
VAR_IN_OUT
  /// Robot assignment of function
  AxesGroup : AxesGroup;
END_VAR

VAR 
  /// internal index
 _idx                       : DINT;
  /// internal sequence index
 _seqIdx                    : DINT;
  /// internal fragment index
 _fragIdx                   : DINT;
  /// internal register index
 _regIdx                    : DINT;
  /// internal execution order list index
 _listIdx                   : DINT := 1;
  /// internal payload pointer
 _payLoadPtr                : DWORD;
  /// internal fragment action
 _fragmentAction            : FragmentAction;
  /// internal fragment action as string
 _fragmentActionString      : STRING;
  /// maximount amount of bytes per sequence
  SEQUENCE_MAX_PAYLOAD_SIZE : UDINT;
END_VAR
                  // ST-FIX F63: the data of a telegram sequence is cleared in AxesGroupToTelegramSequence only
// when it gets a new Seq number; a sequence that is not acknowledged yet is sent unchanged
  
AxesGroupToTelegramHeader        (AxesGroup := AxesGroup);
AxesGroupToTelegramCyclic        (AxesGroup := AxesGroup);
AxesGroupToTelegramCyclicOptional(AxesGroup := AxesGroup);
AxesGroupToTelegramSequence      (AxesGroup := AxesGroup);
AxesGroupToTelegramFooter        (AxesGroup := AxesGroup);
AxesGroupToTelegramLogging       (AxesGroup := AxesGroup);
                
                
END_METHOD

METHOD PRIVATE AxesGroupToTelegramCyclic : DINT
VAR_IN_OUT
  /// Robot assignment of function
  AxesGroup : AxesGroup;
END_VAR
                  IF (AxesGroup.Cyclic.PlcToRob.ToolNo = -1 )
THEN
  Telegram.PlcToRob.Cyclic.ToolNo  := 16#FF;
ELSE
  Telegram.PlcToRob.Cyclic.ToolNo  := INT_TO_BYTE(AxesGroup.Cyclic.PlcToRob.ToolNo); 
END_IF

IF (AxesGroup.Cyclic.PlcToRob.FrameNo = -1 )
THEN
  Telegram.PlcToRob.Cyclic.FrameNo  := 16#FF;
ELSE
  Telegram.PlcToRob.Cyclic.FrameNo  := INT_TO_BYTE(AxesGroup.Cyclic.PlcToRob.FrameNo); 
END_IF
                
END_METHOD

METHOD PRIVATE AxesGroupToTelegramCyclicOptional : DINT
VAR_IN_OUT
  /// Robot assignment of function
  AxesGroup : AxesGroup;
END_VAR
                  // AxesGroup.CyclicOptional.PlcToRob.SubProgramData {{{
IF (AxesGroup.CyclicOptional.PlcToRob.SubProgramData.Active)
THEN
  Telegram.PlcToRob.CyclicOptional.SubProgramData.Data := AxesGroup.CyclicOptional.PlcToRob.SubProgramData.Data; 
END_IF
// }}}

// AxesGroup.CyclicOptional.PlcToRob.CartesianPosition  {{{  
IF (AxesGroup.CyclicOptional.PlcToRob.CartesianPosition.Active)
THEN
  Telegram.PlcToRob.CyclicOptional.CartesianPosition.X           :=                  AxesGroup.CyclicOptional.PlcToRob.CartesianPosition.X;  
  Telegram.PlcToRob.CyclicOptional.CartesianPosition.Y           :=                  AxesGroup.CyclicOptional.PlcToRob.CartesianPosition.Y;  
  Telegram.PlcToRob.CyclicOptional.CartesianPosition.Z           :=                  AxesGroup.CyclicOptional.PlcToRob.CartesianPosition.Z;
  Telegram.PlcToRob.CyclicOptional.CartesianPosition.Rx          :=                  AxesGroup.CyclicOptional.PlcToRob.CartesianPosition.Rx;  
  Telegram.PlcToRob.CyclicOptional.CartesianPosition.Ry          :=                  AxesGroup.CyclicOptional.PlcToRob.CartesianPosition.Ry;  
  Telegram.PlcToRob.CyclicOptional.CartesianPosition.Rz          :=                  AxesGroup.CyclicOptional.PlcToRob.CartesianPosition.Rz;
  Telegram.PlcToRob.CyclicOptional.CartesianPosition.Turns_J2_J1 := CombineHalfSints(AxesGroup.CyclicOptional.PlcToRob.CartesianPosition.TurnNumber.J2Turns, 
                                                                                     AxesGroup.CyclicOptional.PlcToRob.CartesianPosition.TurnNumber.J1Turns);
  Telegram.PlcToRob.CyclicOptional.CartesianPosition.Turns_J4_J3 := CombineHalfSints(AxesGroup.CyclicOptional.PlcToRob.CartesianPosition.TurnNumber.J4Turns, 
                                                                                     AxesGroup.CyclicOptional.PlcToRob.CartesianPosition.TurnNumber.J3Turns);
  Telegram.PlcToRob.CyclicOptional.CartesianPosition.Turns_J6_J5 := CombineHalfSints(AxesGroup.CyclicOptional.PlcToRob.CartesianPosition.TurnNumber.J6Turns, 
                                                                                     AxesGroup.CyclicOptional.PlcToRob.CartesianPosition.TurnNumber.J5Turns);
  // ST-FIX F60: sign + magnitude (spec 5.5.4.4)
  IF ( AxesGroup.CyclicOptional.PlcToRob.CartesianPosition.TurnNumber.E1Turns < 0 )
  THEN
    Telegram.PlcToRob.CyclicOptional.CartesianPosition.Turns_E1 := (INT_TO_BYTE(-SINT_TO_INT(AxesGroup.CyclicOptional.PlcToRob.CartesianPosition.TurnNumber.E1Turns)) AND 16#7F) OR 16#80;
  ELSE
    Telegram.PlcToRob.CyclicOptional.CartesianPosition.Turns_E1 := SINT_TO_BYTE(AxesGroup.CyclicOptional.PlcToRob.CartesianPosition.TurnNumber.E1Turns) AND 16#7F;
  END_IF
END_IF  
// }}}
  
// AxesGroup.CyclicOptional.PlcToRob.CartesianPositionExt {{{ 
IF ( AxesGroup.CyclicOptional.PlcToRob.CartesianPositionExt.Active) 
THEN
  Telegram.PlcToRob.CyclicOptional.CartesianPositionExt.E2 := AxesGroup.CyclicOptional.PlcToRob.CartesianPositionExt.E2;  
  Telegram.PlcToRob.CyclicOptional.CartesianPositionExt.E3 := AxesGroup.CyclicOptional.PlcToRob.CartesianPositionExt.E3;  
  Telegram.PlcToRob.CyclicOptional.CartesianPositionExt.E4 := AxesGroup.CyclicOptional.PlcToRob.CartesianPositionExt.E4;  
  Telegram.PlcToRob.CyclicOptional.CartesianPositionExt.E5 := AxesGroup.CyclicOptional.PlcToRob.CartesianPositionExt.E5;  
  Telegram.PlcToRob.CyclicOptional.CartesianPositionExt.E6 := AxesGroup.CyclicOptional.PlcToRob.CartesianPositionExt.E6;  
END_IF
// }}}

// AxesGroup.CyclicOptional.PlcToRob.JointPosition {{{
IF ( AxesGroup.CyclicOptional.PlcToRob.JointPosition.Active) 
THEN
  Telegram.PlcToRob.CyclicOptional.JointPosition.J1 := AxesGroup.CyclicOptional.PlcToRob.JointPosition.J1;
  Telegram.PlcToRob.CyclicOptional.JointPosition.J2 := AxesGroup.CyclicOptional.PlcToRob.JointPosition.J2;
  Telegram.PlcToRob.CyclicOptional.JointPosition.J3 := AxesGroup.CyclicOptional.PlcToRob.JointPosition.J3;
  Telegram.PlcToRob.CyclicOptional.JointPosition.J4 := AxesGroup.CyclicOptional.PlcToRob.JointPosition.J4;
  Telegram.PlcToRob.CyclicOptional.JointPosition.J5 := AxesGroup.CyclicOptional.PlcToRob.JointPosition.J5;
  Telegram.PlcToRob.CyclicOptional.JointPosition.J6 := AxesGroup.CyclicOptional.PlcToRob.JointPosition.J6;
  Telegram.PlcToRob.CyclicOptional.JointPosition.E1 := AxesGroup.CyclicOptional.PlcToRob.JointPosition.E1;
END_IF
// }}}

// AxesGroup.CyclicOptional.PlcToRob.JointPositionExt {{{
IF ( AxesGroup.CyclicOptional.PlcToRob.JointPositionExt.Active) 
THEN
  Telegram.PlcToRob.CyclicOptional.JointPositionExt.E2 := AxesGroup.CyclicOptional.PlcToRob.JointPositionExt.E2;
  Telegram.PlcToRob.CyclicOptional.JointPositionExt.E3 := AxesGroup.CyclicOptional.PlcToRob.JointPositionExt.E3;  
  Telegram.PlcToRob.CyclicOptional.JointPositionExt.E4 := AxesGroup.CyclicOptional.PlcToRob.JointPositionExt.E4;
  Telegram.PlcToRob.CyclicOptional.JointPositionExt.E5 := AxesGroup.CyclicOptional.PlcToRob.JointPositionExt.E5;
  Telegram.PlcToRob.CyclicOptional.JointPositionExt.E6 := AxesGroup.CyclicOptional.PlcToRob.JointPositionExt.E6;        
END_IF  
// }}}
     
// AxesGroup.CyclicOptional.PlcToRob.Force {{{
IF ( AxesGroup.CyclicOptional.PlcToRob.Force.Active) 
THEN
  Telegram.PlcToRob.CyclicOptional.Force.X  := AxesGroup.CyclicOptional.PlcToRob.Force.X;
  Telegram.PlcToRob.CyclicOptional.Force.Y  := AxesGroup.CyclicOptional.PlcToRob.Force.Y;
  Telegram.PlcToRob.CyclicOptional.Force.Z  := AxesGroup.CyclicOptional.PlcToRob.Force.Z;
  Telegram.PlcToRob.CyclicOptional.Force.Rx := AxesGroup.CyclicOptional.PlcToRob.Force.Rx;
  Telegram.PlcToRob.CyclicOptional.Force.Ry := AxesGroup.CyclicOptional.PlcToRob.Force.Ry;
  Telegram.PlcToRob.CyclicOptional.Force.Rz := AxesGroup.CyclicOptional.PlcToRob.Force.Rz;
END_IF  
// }}}
                    
// AxesGroup.CyclicOptional.PlcToRob.ForceExt {{{
IF ( AxesGroup.CyclicOptional.PlcToRob.ForceExt.Active) 
THEN
  Telegram.PlcToRob.CyclicOptional.ForceExt.E1 := AxesGroup.CyclicOptional.PlcToRob.ForceExt.E1;
  Telegram.PlcToRob.CyclicOptional.ForceExt.E2 := AxesGroup.CyclicOptional.PlcToRob.ForceExt.E2;
  Telegram.PlcToRob.CyclicOptional.ForceExt.E3 := AxesGroup.CyclicOptional.PlcToRob.ForceExt.E3;
  Telegram.PlcToRob.CyclicOptional.ForceExt.E4 := AxesGroup.CyclicOptional.PlcToRob.ForceExt.E4;
  Telegram.PlcToRob.CyclicOptional.ForceExt.E5 := AxesGroup.CyclicOptional.PlcToRob.ForceExt.E5;
  Telegram.PlcToRob.CyclicOptional.ForceExt.E6 := AxesGroup.CyclicOptional.PlcToRob.ForceExt.E6;
END_IF                    
// }}}
                
                
END_METHOD

METHOD PRIVATE AxesGroupToTelegramFooter : DINT
VAR_IN_OUT
  /// Robot assignment of function
  AxesGroup : AxesGroup;
END_VAR
                  Telegram.PlcToRob.Footer.LifeSign := GetHalfeByteLo(Telegram.PlcToRob.Header.FastStop_LifeSign);  
                
END_METHOD

METHOD PRIVATE AxesGroupToTelegramHeader : DINT
VAR_IN_OUT
  /// Robot assignment of function
  AxesGroup : AxesGroup;
END_VAR
                  Telegram.PlcToRob.Header.SRCIVersion               := VersionToByte(AxesGroup.Cyclic.PlcToRob.SRCIVersion);
Telegram.PlcToRob.Header.FastStop_LifeSign         := CombineHalfBytes( HalfByteHi := AxesGroup.Cyclic.PlcToRob.FastStop, HalfByteLo := AxesGroup.Cyclic.PlcToRob.LifeSign );
Telegram.PlcToRob.Header.TelegramLengthPlcToRob    := ParCfg.Com.TelegramLengthPlcToRob;
Telegram.PlcToRob.Header.TelegramLengthRobToPlc    := ParCfg.Com.TelegramLengthRobToPlc;
Telegram.PlcToRob.Header.AxesGroupID_Control       := CombineHalfBytes(HalfByteHi := AxesGroup.Cyclic.PlcToRob.AxesGroupID, HalfByteLo := AxesGroup.Cyclic.PlcToRob.Control);
Telegram.PlcToRob.Header.Reserved                  := 0;
Telegram.PlcToRob.Header.TelegramNumberPlcToRob    := PlcOptionalCyclicToUint(AxesGroup.Parameter.Plc.OptionalCyclic);
Telegram.PlcToRob.Header.TelegramNumberRobToPlc    := RobOptionalCyclicToUint(AxesGroup.Parameter.Rob.OptionalCyclic);
Telegram.PlcToRob.Header.ClientDate                := AxesGroup.Cyclic.PlcToRob.ClientDate;
Telegram.PlcToRob.Header.ClientTime                := AxesGroup.Cyclic.PlcToRob.ClientTime;
                
END_METHOD

METHOD PRIVATE AxesGroupToTelegramLogging : DINT
VAR_IN_OUT
  /// Robot assignment of function
  AxesGroup : AxesGroup;
END_VAR

VAR 
  /// internal sequence index
 _seqIdx                    : DINT;
  /// internal fragment index
 _fragIdx                   : DINT;
END_VAR
                  FOR _seqIdx := 0 TO AxesGroup.State.SequenceCountSend
DO
  // check new data ? 
  IF ( AxesGroup.State.NewSEQ[_seqIdx] )
  THEN
    IF ( Telegram.PlcToRob.Sequence[_seqIdx].Header.PayloadLength > 0 ) 
    THEN
      // Create log entry
      CreateLogMessagePara4 ( Timestamp   := SystemTime,
                              MessageType := MessageType.CMD,
                              Severity    := Severity.DEBUG,
                              MessageCode := 0,
                              MessageText := 'SendData: SEQ = {1}, added Sequence [{2}] with PayloadLength = {3}, HeaderLength = {4}',
                              Para1       :=  UINT_TO_STRING(Telegram.PlcToRob.Sequence[_seqIdx].Header.SEQ_ACK),
                              Para2       :=  DINT_TO_STRING(_seqIdx),
                              Para3       :=  UINT_TO_STRING(Telegram.PlcToRob.Sequence[_seqIdx].Header.PayloadLength),
                              Para4       :=  DINT_TO_STRING(SIZEOF(Telegram.PlcToRob.Sequence[_seqIdx].Header)));
    END_IF
    
    FOR _fragIdx := 0 TO AxesGroup.State.FragmentCountSend[_seqIdx]
    DO
      IF ( Telegram.PlcToRob.Sequence[_seqIdx].Fragment[_fragIdx].Header.PayloadLength > 0 )
      THEN
        // Create log entry
        CreateLogMessagePara6 ( Timestamp   := SystemTime,
                                MessageType := MessageType.CMD,
                                Severity    := Severity.DEBUG,
                                MessageCode := 0,
                                MessageText := 'SendData: added Fragment [{1}] with PayloadLength = {2}, HeaderLength = {3}, CmdID <{4}>, Cmd <{5}> Fragment-Action Bits:{6}' ,
                                Para1       := DINT_TO_STRING(_fragIdx),
                                Para2       := UINT_TO_STRING            (Telegram.PlcToRob.Sequence[_seqIdx].Fragment[_fragIdx].Header.PayloadLength),
                                Para3       := DINT_TO_STRING(SIZEOF     (Telegram.PlcToRob.Sequence[_seqIdx].Fragment[_fragIdx].Header)),                                
                                Para4       := UINT_TO_STRING            (Telegram.PlcToRob.Sequence[_seqIdx].Fragment[_fragIdx].Header.CmdID),
                                Para5       := CMD_TYPE_TO_STRING        (Telegram.PlcToRob.Sequence[_seqIdx].Fragment[_fragIdx].Command.Header.CmdType),
                                Para6       := FRAGMENT_ACTION_TO_STRING (Telegram.PlcToRob.Sequence[_seqIdx].Fragment[_fragIdx].Header.FragmentAction)); 

        // Create log entry
        CreateLogMessagePara2 ( Timestamp   := SystemTime,
                                MessageType := MessageType.CMD,
                                Severity    := Severity.DEBUG,
                                MessageCode := 0,
                                MessageText := 'SendData: added Fragment [{1}] will be executed with ExecMode = [{2}]' ,
                                Para1       := DINT_TO_STRING(_fragIdx),
                                Para2       := EXECUTION_MODE_TO_STRING(Telegram.PlcToRob.Sequence[_seqIdx].Fragment[_fragIdx].Command.Header.ExecMode));

      END_IF
    END_FOR
  END_IF
END_FOR
                
END_METHOD

METHOD PRIVATE AxesGroupToTelegramSequence : DINT
VAR_IN_OUT
  /// Robot assignment of function
  AxesGroup : AxesGroup;
END_VAR

VAR 
  /// internal index
 _idx                       : DINT;
  /// internal sequence index
 _seqIdx                    : DINT;
   /// Amount of sequences
 _seqCount                  : DINT;

  /// internal fragment index
 _fragIdx                   : DINT;
  /// internal register index
 _regIdx                    : DINT;
  /// internal execution order list index
 _listIdx                   : DINT := 1;
  /// internal payload pointer
 _payLoadPtr                : DWORD;
  /// internal fragment action
 _fragmentAction            : FragmentAction;
  /// internal fragment action as string
 _fragmentActionString      : STRING;
  /// maximount amount of bytes per sequence
  SEQUENCE_MAX_PAYLOAD_SIZE : UDINT;
  
  /// current length of telegram 
 _telegramLengthCurrent    : UINT;
END_VAR
                  // Check 2nd sequence active ? 
// ST-FIX F67: remaining space for acyclic data at least 1 byte behind the sequence header
IF ( CalculateSequencePayloadMax(AxesGroup := AxesGroup, Direction := ComDirection.PLC_TO_ROB,
                                 Sequence  := SequenceFlagEnum.PRIMARY_SEQUENCE) < 4 + 1 )
THEN
  SetError( ErrorID := RobotLibraryErrorIdEnum.ERR_ACYCLIC_AREA_TO_SMALL_PLC_TO_ROB, Overwrite := FALSE );
  // Create log entry
  CreateLogMessage ( Timestamp   := SystemTime,
                     MessageType := MessageType.CMD,
                     Severity    := Severity.ERROR,
                     MessageCode := ErrorID,
                     MessageText := 'Telegram PLC -> RC: no space left for acyclic data');
  RETURN;
END_IF
IF ( CalculateSequencePayloadMax(AxesGroup := AxesGroup, Direction := ComDirection.ROB_TO_PLC,
                                 Sequence  := SequenceFlagEnum.PRIMARY_SEQUENCE) < 4 + 1 )
THEN
  SetError( ErrorID := RobotLibraryErrorIdEnum.ERR_ACYCLIC_AREA_TO_SMALL_ROB_TO_PLC, Overwrite := FALSE );
  // Create log entry
  CreateLogMessage ( Timestamp   := SystemTime,
                     MessageType := MessageType.CMD,
                     Severity    := Severity.ERROR,
                     MessageCode := ErrorID,
                     MessageText := 'Telegram RC -> PLC: no space left for acyclic data');
  RETURN;
END_IF

IF ( _parCfg.Com.TwoSequences ) // ST-FIX F63: SEQUENCE_MAX_PAYLOAD_SIZE per sequence, see below
THEN
  // inc sequence counter
 _seqCount := _seqCount + 1;
END_IF   


FOR _seqOrderIdx := 0 TO _seqCount
DO
  // ST-FIX F63: fill the sequence with the lower Seq number first (it is processed first)
  IF ( _seqOrderIdx = 0 )
  THEN
    _seqIdx := _seqSendFirst;
  ELSE
    _seqIdx := 1 - _seqSendFirst;
  END_IF
  // set current SEQ / ACk index
  Telegram.PlcToRob.Sequence[_seqIdx].Header.SEQ_ACK := AxesGroup.State.CurrentSEQ[_seqIdx];

  // only update telegram content if a new sequence SEQ is set
  IF ( AxesGroup.State.NewSEQ[_seqIdx] ) 
  THEN
    // only reset counters in case of new telegram to send  
    // ST-FIX F63: each telegram sequence has its own data area (Fig. 5-205) and starts empty
    IF ( _seqIdx = PRIMARY_SEQUENCE )
    THEN
      SEQUENCE_MAX_PAYLOAD_SIZE := CalculateSequencePayloadMax(AxesGroup := AxesGroup,
                                                               Direction := ComDirection.PLC_TO_ROB,
                                                               Sequence  := SequenceFlagEnum.PRIMARY_SEQUENCE);
    ELSE
      SEQUENCE_MAX_PAYLOAD_SIZE := CalculateSequencePayloadMax(AxesGroup := AxesGroup,
                                                               Direction := ComDirection.PLC_TO_ROB,
                                                               Sequence  := SequenceFlagEnum.SECONDARY_SEQUENCE);
    END_IF
    Telegram.PlcToRob.Sequence[_seqIdx].Header.PayloadLength := 0;
    FOR _idx := 0 TO RobotLibraryParameter.FRAGMENT_MAX
    DO
      Telegram.PlcToRob.Sequence[_seqIdx].Fragment[_idx].Header.PayloadLength := 0;
    END_FOR
   _fragIdx := 0;
   _listIdx := 1;
    AxesGroup.State.FragmentCountSend[_seqIdx] := 0;
    
    // calc current telegram payload length
   _telegramLengthCurrent := 4 + Telegram.PlcToRob.Sequence[_seqIdx].Header.PayloadLength; // ST-FIX F63: sequence header + payload
    
    // Bedingung anpassen und TWO_SEQUENCES berücksichtigen
    WHILE ( _telegramLengthCurrent + FRAGMENT_HEADER_SIZE + MIN_PAYLOAD_SIZE <= SEQUENCE_MAX_PAYLOAD_SIZE ) // ST-FIX F63 
    DO
      // Check command in Execution-Order-List available ?
      IF ( AxesGroup.Acyclic.ActiveCommandRegister.ExecutionOrderList[_listIdx] > EMPTY_EOL_ENTRY)
      THEN
        // set current SEQ / ACk index
        Telegram.PlcToRob.Sequence[_seqIdx].Header.SEQ_ACK := AxesGroup.State.CurrentSEQ[_seqIdx];
        
        // get active command register index
       _regIdx := AxesGroup.Acyclic.ActiveCommandRegister.ExecutionOrderList[_listIdx];
    
        // check State of the current ACR entry ?
        IF (( AxesGroup.Acyclic.ActiveCommandRegister.Register[_regIdx].Command[ACTIVE_CMD].State >= BufferStateCmd.CREATED  ) AND
            ( AxesGroup.Acyclic.ActiveCommandRegister.Register[_regIdx].Command[ACTIVE_CMD].State <= BufferStateCmd.SENDING  ))
        THEN
          // add size of fragement header      
          Telegram.PlcToRob.Sequence[_seqIdx].Header.PayloadLength :=
            Telegram.PlcToRob.Sequence[_seqIdx].Header.PayloadLength + SIZEOF(Telegram.PlcToRob.Sequence[_seqIdx].Fragment[_fragIdx].Header); 
            
            
          Telegram.PlcToRob.Sequence[_seqIdx].Fragment[_fragIdx].Header.CmdID          := AxesGroup.Acyclic.ActiveCommandRegister.Register[_regIdx].UniqueID;
          Telegram.PlcToRob.Sequence[_seqIdx].Fragment[_fragIdx].Header.Reserve        := 0;
          Telegram.PlcToRob.Sequence[_seqIdx].Fragment[_fragIdx].Header.FragmentAction := 0; // will be set below
          Telegram.PlcToRob.Sequence[_seqIdx].Fragment[_fragIdx].Header.PayloadPointer := AxesGroup.Acyclic.ActiveCommandRegister.Register[_regIdx].Command[ACTIVE_CMD].PayLoadPtr; 
          
          // The 1st message resets the ACR entry on the server side  
         _fragmentAction.Reset := (( AxesGroup.Acyclic.ActiveCommandRegister.Register[_regIdx].Command[ACTIVE_CMD].State      = BufferStateCmd.CREATED ) AND
                                   ( AxesGroup.Acyclic.ActiveCommandRegister.Register[_regIdx].Command[ACTIVE_CMD].PayLoadPtr = 0                      ));
                                   
          // Update messages must clear the ACR entry on the server side  
         _fragmentAction.Clear := (( AxesGroup.Acyclic.ActiveCommandRegister.Register[_regIdx].Command[ACTIVE_CMD].State      = BufferStateCmd.UPDATE_AVAILABLE  ) AND
                                   ( AxesGroup.Acyclic.ActiveCommandRegister.Register[_regIdx].Command[ACTIVE_CMD].PayLoadPtr = 0                                )); 
    
          
